(* IEC 61131-3 sources: PortalRobot/Portal_robot/Device/application/FB (part 5) *)

(* ---- FB_ROBOT.st ---- *)
FUNCTION_BLOCK FB_ROBOT
VAR_INPUT
	xUsePhysicalGripperFeedback : BOOL;
	xPhysicalGripperIoReady : BOOL;
	stPhysicalGripperFeedback : ST_GRIPPER_STATUS;
	tPhysicalGripperActionTimeout : TIME := T#10S;
	axMagazineExchangeInProgress : ARRAY [1..2] OF BOOL; // Блокировка адресуется только к меняемому магазину
	xTestInitialize : BOOL;
	auiTestGripperContent : ARRAY [1..2] OF UINT;
	auiTestGripperType : ARRAY [1..2] OF UINT;
	uiTestOrientation : UINT;
	xExternalCommandInhibit : BOOL; // Программный экстренный останов запрещает следующую внешнюю команду
	xSimulationAccelerationEnable : BOOL; // Разрешить ускорение виртуальных таймеров только в симуляции
	uiSimulationTimeFactor : UINT := 1; // Коэффициент виртуального времени 1..100

	stMachine_1_Command : ST_ROBOT_COMMAND; // Команда роботу от первого станка
	stMachine_2_Command : ST_ROBOT_COMMAND; // Команда роботу от второго станка
	stMachine_3_Command : ST_ROBOT_COMMAND; // Команда роботу от третьего станка
	stMagazineCommand   : ST_ROBOT_COMMAND; // Команда роботу от магазина
	stCellCommand       : ST_ROBOT_COMMAND; // Команда позиционирования от менеджера ячейки
	uiBlankPayloadType  : UINT; // Тип заготовки из состояния цикла
	uiDetailPayloadType : UINT; // Тип готовой детали из состояния цикла
	stHmiCommand        : ST_ROBOT_COMMAND; // Ручная команда роботу с HMI
	xReset              : BOOL; // Сброс ошибок робота
	xResetCancel        : BOOL; // Stop/Disable отменяет сброс, не меняя обычную политику останова движения
    xMode               : BOOL; // Режим робота: TRUE — Modbus, FALSE — SoftMotion
	xManual      		: BOOL; // 1 - ручной режим работы, 0 - автоматический режим работы
	xGlobalError        : BOOL; // Глобальная ошибка ячейки
	xEquipmentStopRequired : BOOL; // Владелец оборудования требует зависимую ошибку робота
	ResetDependencies : ST_ROBOT_RESET_DEPENDENCIES; // Снимок отдельных владельцев, только внутренний PLC-контракт
	xModbusBusy         : BOOL; // Внешний робот выполняет команду
	xModbusDone         : BOOL; // Внешний робот завершил команду
	xModbusError        : BOOL; // Ошибка обмена или внешнего робота
	stModbusStatus      : ST_ROBOT_MODBUS_STATUS; // Декодированная обратная связь SC-500
	xHmiDrivesEnable    : BOOL; // Исходный запрос HMI на включение приводов
	xHmiDrivesDisable   : BOOL; // Исходный запрос HMI на отключение приводов
	xHmiStop            : BOOL; // Исходный запрос HMI на остановку
	xHmiDrivesEnableAccepted : BOOL; // RunMotion принял запрос включения в исходном состоянии цикла
	xHmiDrivesDisableAccepted : BOOL; // RunMotion принял запрос отключения в исходном состоянии цикла
	xHmiStopAccepted    : BOOL; // RunMotion принял запрос остановки в исходном состоянии цикла
	xHmiDrivesEnableAllowed : BOOL; // Текущее разрешение включения от владельца Motion-слоя
	xHmiDrivesDisableAllowed : BOOL; // Текущее разрешение отключения от владельца Motion-слоя
	xHmiStopAllowed     : BOOL; // Текущее разрешение остановки от владельца Motion-слоя
	xHmiPermit          : BOOL; // Ручные команды HMI разрешены режимом ячейки
	xManualRecoveryAllowed : BOOL; // Разрешить включение приводов в аварийном ручном восстановлении
	xDrivesPowered      : BOOL; // Все три привода включены
	xDrivesOff          : BOOL; // Все три привода и группа фактически отключены
	xDrivesReady        : BOOL; // Все приводы готовы к движению
	xDriveError         : BOOL; // Активна ошибка оси или группы осей
	xMotionBusy         : BOOL; // Одна из осей выполняет движение
	xMotionResetBusy : BOOL; // Последовательность сброса группы и осей ещё выполняется
	tSoftMotionResetTimeout : TIME := T#30S; // Предел одной принятой попытки сброса
	xSingleAxisMotionBusy : BOOL; // Один из FB_AXIS владеет осью; групповое движение запускать нельзя
	xPointCheckActive : BOOL; // Текущая команда принадлежит проверке сохранённой точки
	xTestAbort : BOOL; // Немедленная отмена активной команды виртуального теста
	rPointCheckSpeedPercent : REAL; // Фактическая скорость проверки 0.1..100 %
	lrGroupAccelerationFactor : LREAL := 1.0; // Общий разгон/торможение групповой траектории, 0.01..1.0
	lrGroupJerkFactor : LREAL := 1.0; // Общий jerk групповой траектории, 0.01..1.0
	tModbusStartTimeout : TIME := T#30S; // Ожидание создания транзакции внешним адаптером
	FaultRequest        : ST_ROBOT_FAULT_REQUEST; // Единый контракт диагностической инъекции
	tGripper1OpenTime   : TIME := T#500MS; // Время открытия первого захвата в модели
	tGripper1CloseTime  : TIME := T#500MS; // Время закрытия первого захвата в модели
	tGripper2OpenTime   : TIME := T#500MS; // Время открытия второго захвата в модели
	tGripper2CloseTime  : TIME := T#500MS; // Время закрытия второго захвата в модели
	tGripperChangeTime  : TIME := T#700MS; // Время смены рабочего захвата в модели

    stPoint : ARRAY [0..GVL_POINT.iPointNumber] OF ST_POINT; // Глобальная таблица точек робота

    xSimBlankAvailable : BOOL; // Начальное наличие заготовки в модели захвата

END_VAR
VAR_OUTPUT
	ResetRecovery : ST_ROBOT_RESET_RECOVERY; // Подтверждение принятой попытки для зависимых владельцев
	GripperCommand : ST_GRIPPER_COMMAND; // Команда для страницы физических выходов
	Command       : ST_ROBOT_COMMAND; // Выбранная команда текущего цикла
	ModbusCommand : ST_ROBOT_COMMAND; // Команда внешнему роботу по Modbus
	Status        : ST_ROBOT_STATUS; // Рабочие статусы робота
	Diag          : ST_ROBOT_DIAG; // Состояние автомата и активная команда
	Error         : ST_ROBOT_ERRORS; // Активные и последние ошибки
	GripperDiag   : ST_GRIPPER_DIAG; // Диагностика внутреннего блока захвата
	GripperError  : ST_GRIPPER_ERRORS; // Активные и последние ошибки захвата
	FaultStatus : ST_ROBOT_FAULT_STATUS; // Сводное состояние инжекторов робота
END_VAR
VAR
	fbMotionManager  : FB_MOTION_MANAGER; // Менеджер перемещения по точкам
    fbGripper        : FB_GRIPPER_SIMULATION; // Модель двухпозиционного захвата
	stGripperCommand : ST_GRIPPER_COMMAND; // Команда внутренней модели захвата

    eState        : E_ROBOT_STATE := E_ROBOT_STATE.IDLE; // Текущее состояние автомата робота
    eActiveAction : E_ROBOT_ACTION := E_ROBOT_ACTION.NONE; // Защёлкнутое действие
    eActivePoint  : E_POINT_NAME; // Защёлкнутая целевая точка
	iActiveSlot   : SINT; // Защёлкнутый слот для всей Modbus-транзакции
	uiActiveMagazineId : UINT; // Защёлкнутый магазин для всей Modbus-транзакции
	uiRobotMagazineContext : UINT; // Физический контекст магазина сохраняется между командами
	xEquipmentStopLatched : BOOL; // Робот остановлен именно аварией обслуживаемого оборудования

	xMotionExecute  : BOOL; // Запрос выполнения перемещения
	xGripperExecute : BOOL; // Запрос выполнения действия захвата
	xManualGripperRequest : BOOL; // Ручной захват разрешён независимо от состояния автомата робота
	xManualGripperOverrideExecute : BOOL; // Прямой импульс FB_GRIPPER из ERROR робота
	eManualGripperAction : E_ROBOT_ACTION; // Действие прямого ручного импульса
	xActiveManualGripper : BOOL; // Текущее действие захвата запущено вручную
	xMagazineCommandActive : BOOL; // Активная команда получена от FB_MAGAZINE
	xMagazineTargetInhibit : BOOL; // Команда входит в магазин, который меняет палеты
	rtReset               : R_TRIG; // Фронт команды сброса робота
	rtHmiDrivesEnable     : R_TRIG; // Фронт запроса включения приводов с HMI
	rtHmiDrivesDisable    : R_TRIG; // Фронт запроса отключения приводов с HMI
	rtHmiStop             : R_TRIG; // Фронт запроса остановки с HMI
	xPowerAllowed         : BOOL; // Визуальная доступность кнопки питания приводов
	xStopAllowed          : BOOL; // Визуальная доступность кнопки остановки
	xResetAllowed         : BOOL; // Визуальная доступность кнопки сброса
	xResetAccepted        : BOOL; // Общий сброс принят владельцем робота
	xExternalResetPending : BOOL; // Удерживает асинхронный Reset до подтверждения SC-500
	xExternalResetIssued  : BOOL; // Reset хотя бы один цикл был передан Modbus-адаптеру
	xSoftMotionResetPending : BOOL; // Один Reset ждёт группу, Motion и захват
	dwResetStopOwners : DWORD; // Владельцы, уже присутствовавшие при принятии Reset
	dwResetLiveCauses : DWORD; // Предыдущий снимок удерживаемых причин этой попытки
	dwResetBusySeen : DWORD; // Владельцы, чей асинхронный сброс действительно запускался
	xEquipmentResetFailed : BOOL; // Новая причина/владелец либо неуспешный терминальный сброс
	tonSoftMotionReset : TON; // Принятая попытка не может оставаться вечной
	xModbusCommandStarted : BOOL; // Текущая команда получила собственную активную транзакцию
	tonModbusStartTimeout : TON; // Защита от вечного ожидания приёма команды адаптером
	fbRobotFaultInjector  : FB_ROBOT_FAULT_INJECTOR; // Безопасная недопустимая команда робота
	xRobotFaultAllowed    : BOOL; // Владелец готов проверить тестовую команду
	uiTestBlankPayloadType : UINT;
	uiTestDetailPayloadType : UINT;
	xTestBlankPayloadPending : BOOL;
	xTestDetailPayloadPending : BOOL;

END_VAR

VAR_IN_OUT
    stMotionManager : ST_MOTION_MANAGER; // Данные менеджера движения
    GroupData       : ST_AXIS_GROUP; // Данные группы осей XYZ
    stPointManager  : ST_POINT_MANAGER; // Данные проверки точки
END_VAR

VAR CONSTANT
	ERR_ROBOT_WRONG_ACTION : DWORD := DWORD#16#0000_0001; // Недопустимое действие робота
    ERR_ROBOT_MOTION       : DWORD := DWORD#16#0000_0002; // Ошибка менеджера движения
    ERR_ROBOT_GRIPPER      : DWORD := DWORD#16#0000_0004; // Ошибка захвата
	ERR_ROBOT_MODBUS_COMM  : DWORD := DWORD#16#0000_0008; // Ошибка связи Modbus TCP
	ERR_ROBOT_STOP         : DWORD := DWORD#16#0000_0010; // Остановка команды робота
	ERR_EXTERNAL_ROBOT     : DWORD := DWORD#16#0000_0020; // Контроллер робота сообщил аварию
	WRN_RESET_EXECUTE_ACTIVE : UINT := 1; // Команда робота ещё активна
	WRN_RESET_STOP_ACTIVE    : UINT := 2; // Команда остановки ещё активна
	WRN_RESET_GLOBAL_ERROR   : UINT := 3; // Глобальная ошибка ещё активна
	WRN_RESET_MOTION_ERROR   : UINT := 4; // Ошибка менеджера движения ещё активна
	WRN_RESET_GRIPPER_ERROR  : UINT := 5; // Ошибка захвата ещё активна
	WRN_RESET_MODBUS_ERROR   : UINT := 6; // Ошибка внешнего робота ещё активна
	WRN_HMI_MANUAL_REQUIRED  : UINT := 7; // Ручная команда запрещена режимом ячейки
	WRN_DRIVES_ENABLE_ERROR  : UINT := 8; // Команда приводов отклонена владельцем Motion-слоя
	WRN_STOP_DRIVES_NOT_READY: UINT := 9; // Остановка недоступна при неготовых приводах
	WRN_SIM_ERROR_NOT_ALLOWED: UINT := 11; // Тестовая команда запрещена текущим состоянием
	WRN_RESET_EQUIPMENT_ERROR : UINT := 18; // WARNING через общий канал: зависимый сброс прерван/не завершён
END_VAR

// --- BEGIN IMPLEMENTATION ---

rtHmiDrivesEnable(CLK := xHmiDrivesEnable);
rtHmiDrivesDisable(CLK := xHmiDrivesDisable);
rtHmiStop(CLK := xHmiStop);

xPowerAllowed := ((NOT xDrivesOff) AND xHmiDrivesDisableAllowed)
	OR (xDrivesOff AND xHmiDrivesEnableAllowed);
xStopAllowed := xHmiStopAllowed;

IF (rtHmiDrivesEnable.Q AND NOT xHmiDrivesEnableAccepted)
OR (rtHmiDrivesDisable.Q AND NOT xHmiDrivesDisableAccepted) THEN
	IF NOT xHmiPermit THEN
		Diag.stWarning.uiCode := WRN_HMI_MANUAL_REQUIRED;
	ELSE
		Diag.stWarning.uiCode := WRN_DRIVES_ENABLE_ERROR;
	END_IF;
	Diag.stWarning.udiSequence := Diag.stWarning.udiSequence + UDINT#1;
	IF Diag.stWarning.udiSequence = UDINT#0 THEN
		Diag.stWarning.udiSequence := UDINT#1;
	END_IF;
END_IF;

IF rtHmiStop.Q
AND NOT xHmiStopAccepted THEN
	IF NOT xHmiPermit THEN
		Diag.stWarning.uiCode := WRN_HMI_MANUAL_REQUIRED;
	ELSE
		Diag.stWarning.uiCode := WRN_STOP_DRIVES_NOT_READY;
	END_IF;
	Diag.stWarning.udiSequence := Diag.stWarning.udiSequence + UDINT#1;
	IF Diag.stWarning.udiSequence = UDINT#0 THEN
		Diag.stWarning.udiSequence := UDINT#1;
	END_IF;
END_IF;

// Команды по умолчанию
xMotionExecute := FALSE;
xGripperExecute := FALSE;
xManualGripperRequest := FALSE;
xManualGripperOverrideExecute := FALSE;
xMagazineCommandActive := FALSE;
xMagazineTargetInhibit := FALSE;

Command.xExecute := FALSE;
Command.xStop := FALSE;
Command.xReset := FALSE;
Command.eAction := E_ROBOT_ACTION.NONE;
Command.eSetPoint := E_POINT_NAME.NONE;
Command.iActiveSlot := 0;
Command.uiMagazineId := UINT#0;

ModbusCommand.xExecute := FALSE;
ModbusCommand.xStop := FALSE;
ModbusCommand.xReset := FALSE;
ModbusCommand.eAction := E_ROBOT_ACTION.NONE;
ModbusCommand.eSetPoint := E_POINT_NAME.NONE;
ModbusCommand.iActiveSlot := 0;
ModbusCommand.uiMagazineId := UINT#0;

//Определяем какой режим работы активен
IF NOT xManual THEN
	IF stCellCommand.xExecute OR stCellCommand.xStop THEN
		Command := stCellCommand;
	ELSIF stMachine_1_Command.xExecute OR stMachine_1_Command.xStop THEN
		Command := stMachine_1_Command;
	ELSIF stMachine_2_Command.xExecute OR stMachine_2_Command.xStop THEN
		Command := stMachine_2_Command;
	ELSIF stMachine_3_Command.xExecute OR stMachine_3_Command.xStop THEN
		Command := stMachine_3_Command;
	ELSIF stMagazineCommand.xExecute OR stMagazineCommand.xStop THEN
		Command := stMagazineCommand;
		xMagazineCommandActive := TRUE;
	END_IF;
ELSE
	IF stMagazineCommand.xExecute OR stMagazineCommand.xStop THEN
		Command := stMagazineCommand;
		xMagazineCommandActive := TRUE;
	ELSE
		Command := stHmiCommand;
	END_IF;
END_IF;

// Смена палет блокирует автоматические команды и операции FB_MAGAZINE
// с этим магазином. Ручная точка HMI не зависит от состояния магазина.
IF (NOT xManual OR xMagazineCommandActive)
AND (Command.uiMagazineId >= UINT#1) AND (Command.uiMagazineId <= UINT#2) THEN
	IF axMagazineExchangeInProgress[Command.uiMagazineId] THEN
		IF (Command.eSetPoint = E_POINT_NAME.MAGAZINE_SAFE)
		OR (Command.eSetPoint = E_POINT_NAME.MAGAZINE_CHANGE)
		OR (Command.eSetPoint = E_POINT_NAME.MAGAZINE_IN_SLOT) THEN
			xMagazineTargetInhibit := TRUE;
		END_IF;
	END_IF;
END_IF;

// Abort теста имеет приоритет над любым владельцем, включая ручную подготовку
// сценария, когда команда ячейки обычно не участвует в выборе.
IF xTestAbort THEN
	Command.xExecute := FALSE;
	Command.xStop := TRUE;
END_IF;

// Уже принятую внешним контроллером команду не прерываем. Запрет действует
// только в IDLE, то есть перед началом следующего высокоуровневого действия.
IF xMode
AND xExternalCommandInhibit
AND (eState = E_ROBOT_STATE.IDLE) THEN
	Command.xExecute := FALSE;
END_IF;

IF xMagazineTargetInhibit AND (eState = E_ROBOT_STATE.IDLE) THEN
	Command.xExecute := FALSE;
END_IF;

// Внешний Stop — самостоятельная приоритетная команда. Он должен дойти до
// адаптера и тогда, когда FB_ROBOT уже защёлкнул ERROR после общей остановки.
IF xMode
AND (xHmiStopAccepted
	OR Command.xStop
	OR (xGlobalError AND stModbusStatus.xBusy)) THEN
	ModbusCommand.xStop := TRUE;
END_IF;

// Класс ошибки определяет оборудование-владелец. FB_ROBOT только выполняет
// зависимую реакцию: активное действие останавливает, неподвижный робот сразу
// переводит в ERROR без бессмысленной команды Stop.
IF xEquipmentStopRequired
AND (eState <> E_ROBOT_STATE.ERROR) THEN
	xEquipmentStopLatched := TRUE;
	IF (eState = E_ROBOT_STATE.MOTION)
	OR (eState = E_ROBOT_STATE.GRIPPER)
	OR (eState = E_ROBOT_STATE.MODBUS) THEN
		Command.xStop := TRUE;
	ELSE
		Error.dwErrorActive := Error.dwErrorActive OR ERR_ROBOT_STOP;
		eState := E_ROBOT_STATE.ERROR;
	END_IF;
END_IF;

// RunRobot уже выполнил все PLC-проверки и передал Execute только принятой
// ручной команде. Захват остаётся независимым от состояния осей и робота.
IF xManual AND stHmiCommand.xExecute THEN
	CASE stHmiCommand.eAction OF
		E_ROBOT_ACTION.UNCLAMP_1,
		E_ROBOT_ACTION.CLAMP_1,
		E_ROBOT_ACTION.UNCLAMP_2,
		E_ROBOT_ACTION.CLAMP_2,
		E_ROBOT_ACTION.ROTATE_TO_BLANK,
		E_ROBOT_ACTION.ROTATE_TO_DETAIL:
			xManualGripperRequest := TRUE;
	END_CASE;
END_IF;

// Готовность сброса рассчитывается после выбора актуального владельца команды.
// Ошибки вложенных FB считаются сбрасываемыми только после снятия удерживаемого
// источника и публикации их собственного xResetAllowed.
rtReset(CLK := xReset);
xResetAllowed := xHmiPermit AND NOT xResetCancel
	AND NOT xTestAbort AND NOT xHmiStop AND NOT xHmiStopAccepted
	AND NOT xSoftMotionResetPending
	AND NOT xExternalResetPending
	AND (NOT xMode OR NOT stModbusStatus.xResetBusy)
	AND (NOT xGlobalError OR xManualRecoveryAllowed)
	AND NOT Command.xExecute
	AND NOT Command.xStop
	AND NOT xMotionBusy
	AND (NOT xMode OR stModbusStatus.xCommunicationAlive)
	AND (xDriveError
		OR (eState = E_ROBOT_STATE.ERROR)
		OR (NOT xMode AND stMotionManager.Status.xError)
		OR (NOT xMode AND fbGripper.Status.xError)
		OR (xMode AND xModbusError))
	AND (xMode OR NOT stMotionManager.Status.xError
		OR FaultStatus.stPoint.xResetAllowed)
	AND (xMode OR NOT fbGripper.Status.xError
		OR FaultStatus.stGripper.xResetAllowed);
xResetAccepted := rtReset.Q AND xResetAllowed;
IF xResetAccepted THEN
	ResetRecovery.udiAttempt := ResetRecovery.udiAttempt + UDINT#1;
	IF ResetRecovery.udiAttempt = UDINT#0 THEN ResetRecovery.udiAttempt := UDINT#1; END_IF;
	dwResetStopOwners := ResetDependencies.dwStopOwners;
	dwResetLiveCauses := ResetDependencies.dwLiveCauses;
	dwResetBusySeen := ResetDependencies.dwResetBusy;
END_IF;
xEquipmentResetFailed := FALSE;
IF (xSoftMotionResetPending OR xExternalResetPending) AND NOT xResetAccepted THEN
	// Нового владельца или повторный фронт физической причины нельзя принять
	// за хвост старого сброса. Падение Busy само по себе успехом не является.
	xEquipmentResetFailed := ((ResetDependencies.dwStopOwners AND NOT dwResetStopOwners) <> DWORD#0)
		OR ((ResetDependencies.dwLiveCauses AND NOT dwResetLiveCauses) <> DWORD#0)
		OR ((dwResetBusySeen AND NOT ResetDependencies.dwResetBusy
			AND ResetDependencies.dwStopOwners) <> DWORD#0);
	dwResetLiveCauses := ResetDependencies.dwLiveCauses;
	dwResetBusySeen := dwResetBusySeen OR ResetDependencies.dwResetBusy;
END_IF;
// Общий Reset запускает Motion-сброс раньше FB_ROBOT. Если группа была в
// ErrorStop, одноцикловый импульс уже закончится к моменту её восстановления;
// защёлкиваем намерение оператора до исчезновения первичной Motion-ошибки.
IF xMode THEN
	xSoftMotionResetPending := FALSE;
ELSIF xResetAccepted
AND (eState = E_ROBOT_STATE.ERROR) THEN
	xSoftMotionResetPending := TRUE;
END_IF;
IF xMode AND xResetAccepted THEN
	xExternalResetPending := TRUE;
	xExternalResetIssued := FALSE;
ELSIF NOT xMode THEN
	xExternalResetPending := FALSE;
	xExternalResetIssued := FALSE;
END_IF;

tonSoftMotionReset(IN := xSoftMotionResetPending OR xExternalResetPending, PT := tSoftMotionResetTimeout);
IF xSoftMotionResetPending AND NOT xResetAccepted
AND (tonSoftMotionReset.Q
	OR xEquipmentResetFailed OR xResetCancel
	OR xTestAbort OR NOT xHmiPermit OR Command.xExecute OR Command.xStop OR xHmiStop OR xHmiStopAccepted
	OR (xGlobalError AND NOT xManualRecoveryAllowed)
	OR (xDriveError AND NOT xMotionResetBusy)
	OR (fbGripper.Status.xError AND NOT FaultStatus.stGripper.xResetAllowed)
	OR (stMotionManager.Status.xError AND NOT FaultStatus.stPoint.xResetAllowed)) THEN
	xSoftMotionResetPending := FALSE;
	IF xEquipmentResetFailed OR (tonSoftMotionReset.Q AND xEquipmentStopRequired) THEN
		Diag.stWarning.uiCode := WRN_RESET_EQUIPMENT_ERROR;
	ELSIF fbGripper.Status.xError THEN
		Diag.stWarning.uiCode := WRN_RESET_GRIPPER_ERROR;
	ELSE
		Diag.stWarning.uiCode := WRN_RESET_MOTION_ERROR;
	END_IF;
	Diag.stWarning.udiSequence := Diag.stWarning.udiSequence + UDINT#1;
	IF Diag.stWarning.udiSequence = UDINT#0 THEN Diag.stWarning.udiSequence := UDINT#1; END_IF;
END_IF;

// После неуспешной попытки адаптер публикует явный результат. Снимаем уровень,
// чтобы следующее осознанное нажатие Reset снова дошло до его R_TRIG.
IF xExternalResetPending AND xExternalResetIssued AND NOT xResetAccepted
AND (stModbusStatus.xResetFailed OR NOT stModbusStatus.xCommunicationAlive
	OR tonSoftMotionReset.Q OR xEquipmentResetFailed OR xResetCancel
	OR xTestAbort OR Command.xStop OR xHmiStop OR xHmiStopAccepted OR NOT xHmiPermit
	OR (xGlobalError AND NOT xManualRecoveryAllowed)) THEN
	xExternalResetPending := FALSE;
	xExternalResetIssued := FALSE;
	IF xEquipmentResetFailed OR (tonSoftMotionReset.Q AND xEquipmentStopRequired) THEN
		Diag.stWarning.uiCode := WRN_RESET_EQUIPMENT_ERROR;
	ELSE
		Diag.stWarning.uiCode := WRN_RESET_MODBUS_ERROR;
	END_IF;
	Diag.stWarning.udiSequence := Diag.stWarning.udiSequence + UDINT#1;
	IF Diag.stWarning.udiSequence = UDINT#0 THEN Diag.stWarning.udiSequence := UDINT#1; END_IF;
END_IF;

// Недопустимое действие проверяется в IDLE до запуска Motion или захвата.
xRobotFaultAllowed := (eState = E_ROBOT_STATE.IDLE)
	AND NOT Command.xExecute
	AND NOT Command.xStop
	AND NOT xMode
	AND NOT xGlobalError
	AND NOT xDriveError
	AND (Error.dwErrorActive = DWORD#0)
	AND NOT stMotionManager.Status.xError
	AND NOT fbGripper.Status.xError;

fbRobotFaultInjector(
	Request := FaultRequest,
	xOwnerAllowed := xRobotFaultAllowed
);
FaultStatus.stRobot := fbRobotFaultInjector.Status;

IF fbRobotFaultInjector.Status.xRejected THEN
	Diag.stWarning.uiCode := WRN_SIM_ERROR_NOT_ALLOWED;
	Diag.stWarning.udiSequence := Diag.stWarning.udiSequence + UDINT#1;
	IF Diag.stWarning.udiSequence = UDINT#0 THEN
		Diag.stWarning.udiSequence := UDINT#1;
	END_IF;
END_IF;

IF fbRobotFaultInjector.xWrongAction THEN
	Command.xExecute := TRUE;
	Command.xStop := FALSE;
	Command.eAction := E_ROBOT_ACTION.NONE;
	Command.eSetPoint := E_POINT_NAME.NONE;
END_IF;

Command.xReset := xResetAccepted;

IF rtReset.Q
AND ((eState = E_ROBOT_STATE.ERROR) OR xDriveError)
AND NOT xResetAccepted THEN
	IF NOT xHmiPermit THEN
		Diag.stWarning.uiCode := WRN_HMI_MANUAL_REQUIRED;
	ELSIF eState <> E_ROBOT_STATE.ERROR THEN
		// Ошибку Motion-слоя сбрасывают оси и группа тем же общим импульсом.
		Diag.stWarning.uiCode := UINT#0;
    ELSIF Command.xExecute THEN
        Diag.stWarning.uiCode := WRN_RESET_EXECUTE_ACTIVE;
    ELSIF Command.xStop THEN
        Diag.stWarning.uiCode := WRN_RESET_STOP_ACTIVE;
    ELSIF xGlobalError AND NOT xManualRecoveryAllowed THEN
        Diag.stWarning.uiCode := WRN_RESET_GLOBAL_ERROR;
    ELSIF stMotionManager.Status.xError
	OR (NOT xMode AND xDriveError) THEN
        Diag.stWarning.uiCode := WRN_RESET_MOTION_ERROR;
    ELSIF fbGripper.Status.xError THEN
        Diag.stWarning.uiCode := WRN_RESET_GRIPPER_ERROR;
    ELSIF xModbusError THEN
        Diag.stWarning.uiCode := WRN_RESET_MODBUS_ERROR;
    ELSE
        Diag.stWarning.uiCode := UINT#0;
    END_IF;

    IF Diag.stWarning.uiCode <> UINT#0 THEN
        Diag.stWarning.udiSequence := Diag.stWarning.udiSequence + UDINT#1;
        IF Diag.stWarning.udiSequence = UDINT#0 THEN
            Diag.stWarning.udiSequence := UDINT#1;
        END_IF;
    END_IF;
END_IF;

// =====================================================
// Автомат FB_ROBOT
// =====================================================

// Таймаут исполнения принадлежит FB_ROBOT_MODBUS, но до создания активной
// транзакции его TON ещё не работает. Отдельно ограничиваем фазу ожидания Busy.
tonModbusStartTimeout(
	IN := xMode
		AND (eState = E_ROBOT_STATE.MODBUS)
		AND NOT xModbusCommandStarted,
	PT := tModbusStartTimeout
);

// Ошибка оси или группы является первопричиной в Motion-слое и отдельной
// каскадной ошибкой робота для его публичного статуса и журнала.
IF NOT xMode AND xDriveError THEN
	Error.dwErrorActive := Error.dwErrorActive OR ERR_ROBOT_MOTION;
	eState := E_ROBOT_STATE.ERROR;
ELSIF NOT xMode AND stMotionManager.Status.xError THEN
	// Отмена задания при ручном I/O не скрывает аварию вложенного владельца.
	Error.dwErrorActive := Error.dwErrorActive OR ERR_ROBOT_MOTION;
	eState := E_ROBOT_STATE.ERROR;
ELSIF NOT xMode AND fbGripper.Status.xError THEN
	Error.dwErrorActive := Error.dwErrorActive OR ERR_ROBOT_GRIPPER;
	eState := E_ROBOT_STATE.ERROR;
ELSIF xMode AND xModbusError THEN
	IF stModbusStatus.xRobotAlarm THEN
		Error.dwErrorActive := Error.dwErrorActive OR ERR_EXTERNAL_ROBOT;
	ELSE
		Error.dwErrorActive := Error.dwErrorActive OR ERR_ROBOT_MODBUS_COMM;
	END_IF;
	eState := E_ROBOT_STATE.ERROR;
END_IF;

CASE eState OF

    E_ROBOT_STATE.IDLE:

        Status.xBusy := FALSE;
        Status.xDone := FALSE;
        Status.xError := FALSE;

        IF Command.xExecute THEN
            eActiveAction := Command.eAction;
            eActivePoint := Command.eSetPoint;
			iActiveSlot := Command.iActiveSlot;
			uiActiveMagazineId := Command.uiMagazineId;
			IF (Command.uiMagazineId >= UINT#1)
			AND (Command.uiMagazineId <= UINT#2)
			AND (Command.eAction = E_ROBOT_ACTION.MOVE_TO_POINT)
			AND ((Command.eSetPoint = E_POINT_NAME.MAGAZINE_IN_SLOT)
				OR (Command.eSetPoint = E_POINT_NAME.MAGAZINE_CHANGE)) THEN
				uiRobotMagazineContext := Command.uiMagazineId;
			END_IF;

            IF xMode THEN
				xModbusCommandStarted := FALSE;
				eState := E_ROBOT_STATE.MODBUS;

            ELSE
                CASE Command.eAction OF

                    E_ROBOT_ACTION.MOVE_TO_POINT:
                        // CODESYS переводит группу в ошибку, если GroupMoving
                        // запускается при активном single-axis FB. Команда
                        // остаётся в IDLE до освобождения всех FB_AXIS.
                        IF xDrivesReady AND NOT xMotionBusy THEN
                            eState := E_ROBOT_STATE.MOTION;
                        END_IF;

                    E_ROBOT_ACTION.UNCLAMP_1,
                    E_ROBOT_ACTION.CLAMP_1,
                    E_ROBOT_ACTION.UNCLAMP_2,
                    E_ROBOT_ACTION.CLAMP_2,
                    E_ROBOT_ACTION.ROTATE_TO_BLANK,
                    E_ROBOT_ACTION.ROTATE_TO_DETAIL:
						xActiveManualGripper := xManualGripperRequest;
                        eState := E_ROBOT_STATE.GRIPPER;

                ELSE
                    Error.dwErrorActive :=
                        Error.dwErrorActive OR ERR_ROBOT_WRONG_ACTION;

                    eState := E_ROBOT_STATE.ERROR;
                END_CASE;
            END_IF;
        END_IF;

    E_ROBOT_STATE.MOTION:

        Status.xBusy := TRUE;
        xMotionExecute := NOT xSingleAxisMotionBusy;

		IF xHmiStopAccepted OR Command.xStop THEN
			// Операторский Stop отменяет действие штатно. Stop от оборудования
			// дополнительно защёлкивает зависимую ошибку робота.
            xMotionExecute := FALSE;
            Status.xBusy := FALSE;
            Status.xDone := FALSE;
            eActiveAction := E_ROBOT_ACTION.NONE;
            eActivePoint := E_POINT_NAME.NONE;
			IF xEquipmentStopRequired THEN
				Error.dwErrorActive := Error.dwErrorActive OR ERR_ROBOT_STOP;
				eState := E_ROBOT_STATE.ERROR;
			ELSE
				eState := E_ROBOT_STATE.IDLE;
			END_IF;

        ELSIF xGlobalError THEN
            Error.dwErrorActive := Error.dwErrorActive OR ERR_ROBOT_STOP;
            eState := E_ROBOT_STATE.ERROR;

        ELSIF stMotionManager.Status.xError THEN
            Error.dwErrorActive := Error.dwErrorActive OR ERR_ROBOT_MOTION;
            eState := E_ROBOT_STATE.ERROR;

		ELSIF stMotionManager.Status.xDone THEN
			IF (eActiveAction = E_ROBOT_ACTION.MOVE_TO_POINT)
			AND (eActivePoint <> E_POINT_NAME.MAGAZINE_IN_SLOT)
			AND (eActivePoint <> E_POINT_NAME.MAGAZINE_CHANGE) THEN
				uiRobotMagazineContext := UINT#0;
			END_IF;
            eState := E_ROBOT_STATE.DONE;
        END_IF;

	E_ROBOT_STATE.GRIPPER:

        Status.xBusy := TRUE;
        xGripperExecute := TRUE;

		IF xTestAbort THEN
			xGripperExecute := FALSE;
			Status.xBusy := FALSE;
			Status.xDone := FALSE;
			xActiveManualGripper := FALSE;
			eActiveAction := E_ROBOT_ACTION.NONE;
			eActivePoint := E_POINT_NAME.NONE;
			eState := E_ROBOT_STATE.IDLE;

		ELSIF xEquipmentStopRequired THEN
			xGripperExecute := FALSE;
			Error.dwErrorActive := Error.dwErrorActive OR ERR_ROBOT_STOP;
			eState := E_ROBOT_STATE.ERROR;

		ELSIF xGlobalError AND NOT xActiveManualGripper THEN
            Error.dwErrorActive := Error.dwErrorActive OR ERR_ROBOT_STOP;
            eState := E_ROBOT_STATE.ERROR;

        ELSIF fbGripper.Status.xError THEN
            Error.dwErrorActive := Error.dwErrorActive OR ERR_ROBOT_GRIPPER;
            eState := E_ROBOT_STATE.ERROR;

        ELSIF fbGripper.Status.xDone THEN
			xActiveManualGripper := FALSE;
            eState := E_ROBOT_STATE.DONE;
        END_IF;

	E_ROBOT_STATE.DONE:

        Status.xBusy := FALSE;
        Status.xDone := TRUE;

        IF NOT xMode THEN
        CASE eActiveAction OF

            E_ROBOT_ACTION.MOVE_TO_POINT:
                xMotionExecute := TRUE;

            E_ROBOT_ACTION.UNCLAMP_1,
            E_ROBOT_ACTION.CLAMP_1,
            E_ROBOT_ACTION.UNCLAMP_2,
            E_ROBOT_ACTION.CLAMP_2,
            E_ROBOT_ACTION.ROTATE_TO_BLANK,
            E_ROBOT_ACTION.ROTATE_TO_DETAIL:
                xGripperExecute := TRUE;

        END_CASE;
        END_IF;

		IF NOT Command.xExecute THEN
			// Владелец уже снял Execute: в этом же цикле погасить запрос
			// вложенному FB до очистки action/point. Иначе при быстром
			// SoftMotion движении один скан уходил как Execute=TRUE + point=NONE,
			// а FB_MOTION_MANAGER закономерно валил нулевую точку.
			xMotionExecute := FALSE;
			xGripperExecute := FALSE;
            Status.xDone := FALSE;
			xModbusCommandStarted := FALSE;
            eActiveAction := E_ROBOT_ACTION.NONE;
			eActivePoint := E_POINT_NAME.NONE;
			iActiveSlot := SINT#0;
			uiActiveMagazineId := UINT#0;
			eState := E_ROBOT_STATE.IDLE;
        END_IF;

	E_ROBOT_STATE.MODBUS:
		Status.xBusy := TRUE;
		// Execute — импульс от владельца команды. Адаптер Modbus может
		// быть занят FC03/FC16 дольше этого импульса. Поэтому до терминального
		// ответа передаём защёлкнутые action/point/slot, а не уже снятый Command.
		ModbusCommand.xExecute := TRUE;
		ModbusCommand.eAction := eActiveAction;
		ModbusCommand.eSetPoint := eActivePoint;
		ModbusCommand.iActiveSlot := iActiveSlot;
		ModbusCommand.uiMagazineId := uiActiveMagazineId;
		IF xModbusBusy THEN
			xModbusCommandStarted := TRUE;
		END_IF;

		IF xTestAbort THEN
			ModbusCommand.xStop := TRUE;
			IF NOT stModbusStatus.xBusy THEN
				Status.xBusy := FALSE;
				Status.xDone := FALSE;
				xModbusCommandStarted := FALSE;
				eActiveAction := E_ROBOT_ACTION.NONE;
				eActivePoint := E_POINT_NAME.NONE;
				iActiveSlot := SINT#0;
				uiActiveMagazineId := UINT#0;
				eState := E_ROBOT_STATE.IDLE;
			END_IF;
		ELSIF Command.xStop OR xHmiStopAccepted OR xGlobalError THEN
			ModbusCommand.xStop := TRUE;
			Error.dwErrorActive := Error.dwErrorActive OR ERR_ROBOT_STOP;
			eState := E_ROBOT_STATE.ERROR;
		ELSIF xModbusError THEN
			IF stModbusStatus.xRobotAlarm THEN
				Error.dwErrorActive := Error.dwErrorActive OR ERR_EXTERNAL_ROBOT;
			ELSE
				Error.dwErrorActive := Error.dwErrorActive OR ERR_ROBOT_MODBUS_COMM;
			END_IF;
			eState := E_ROBOT_STATE.ERROR;
		ELSIF tonModbusStartTimeout.Q THEN
			// Адаптер не создал собственную транзакцию: не оставляем публичный
			// xBusy висеть бесконечно без CommandSeq и физического движения.
			ModbusCommand.xExecute := FALSE;
			Error.dwErrorActive := Error.dwErrorActive OR ERR_ROBOT_MODBUS_COMM;
			eState := E_ROBOT_STATE.ERROR;
		ELSIF xModbusCommandStarted AND xModbusDone THEN
			IF (eActiveAction = E_ROBOT_ACTION.MOVE_TO_POINT)
			AND (eActivePoint <> E_POINT_NAME.MAGAZINE_IN_SLOT)
			AND (eActivePoint <> E_POINT_NAME.MAGAZINE_CHANGE) THEN
				uiRobotMagazineContext := UINT#0;
			END_IF;
			eState := E_ROBOT_STATE.DONE;
		END_IF;

    E_ROBOT_STATE.ERROR:

        Status.xBusy := FALSE;
        Status.xDone := FALSE;
        Status.xError := TRUE;

		// Ошибка координатного робота не блокирует независимый ручной захват.
		// Собственная ошибка FB_GRIPPER по-прежнему требует штатного сброса.
		IF NOT xMode AND xManualGripperRequest AND NOT fbGripper.Status.xError THEN
			xManualGripperOverrideExecute := TRUE;
			eManualGripperAction := stHmiCommand.eAction;
		END_IF;

		// В Modbus-режиме входной Reset только защёлкивает запрос для адаптера.
		// Локальную ошибку можно снять лишь после подтверждённого исчезновения
		// внешней аварии; иначе xExternalResetPending очистится до записи 1004.
		IF ((NOT xMode AND (xResetAccepted OR xSoftMotionResetPending))
			OR (xMode
				AND xExternalResetPending
				AND xExternalResetIssued
				AND stModbusStatus.xResetDone
				AND NOT xModbusError
				AND NOT stModbusStatus.xBusy
				AND (stModbusStatus.uiExecutionState =
					TO_UINT(E_ROBOT_MODBUS_EXECUTION_STATE.IDLE))))
        AND NOT Command.xExecute
        AND NOT Command.xStop
        AND NOT xEquipmentStopRequired
        AND (NOT xGlobalError OR xManualRecoveryAllowed)
		AND (xMode OR NOT stMotionManager.Status.xError)
		AND (xMode OR NOT xDriveError)
		AND (xMode OR NOT xMotionResetBusy)
		AND (xMode OR NOT fbGripper.Status.xError)
		AND (NOT xMode OR stModbusStatus.xCommunicationAlive) THEN

			Error.dwErrorLast := Error.dwErrorActive;
			Error.dwErrorActive := DWORD#0;
            Status.xError := FALSE;
			xExternalResetPending := FALSE;
			xExternalResetIssued := FALSE;
			xSoftMotionResetPending := FALSE;
			xModbusCommandStarted := FALSE;
			xActiveManualGripper := FALSE;
			xEquipmentStopLatched := FALSE;
            eActiveAction := E_ROBOT_ACTION.NONE;
			eActivePoint := E_POINT_NAME.NONE;
			iActiveSlot := SINT#0;
			uiActiveMagazineId := UINT#0;
			eState := E_ROBOT_STATE.IDLE;
        END_IF;

END_CASE;

IF xMode AND xExternalResetPending THEN
	ModbusCommand.xReset := TRUE;
	xExternalResetIssued := TRUE;
END_IF;

// =====================================================
// Формирование команды FB_MOTION_MANAGER
// =====================================================

stMotionManager.Command.xExecute := NOT xMode AND xMotionExecute;
stMotionManager.Command.eTargetPoint := eActivePoint;
stMotionManager.Command.xReset := NOT xMode AND xResetAccepted;
stMotionManager.Command.xStop := NOT xMode AND (xHmiStopAccepted OR Command.xStop);
stMotionManager.Command.xGlobalError :=
    (NOT xMode AND xGlobalError AND NOT xManualRecoveryAllowed);

// =====================================================
// Вызов FB_MOTION_MANAGER
// =====================================================

fbMotionManager(
    stPoint := stPoint,
    xReset := NOT xMode AND xResetAccepted,
	FaultRequest := FaultRequest.stPoint,
	xSpeedFactorOverride := xPointCheckActive,
	lrSpeedFactorOverride := REAL_TO_LREAL(rPointCheckSpeedPercent) / 100.0,
	lrAccelerationFactor := lrGroupAccelerationFactor,
	lrJerkFactor := lrGroupJerkFactor,
    stMotionManager := stMotionManager,
    GroupData := GroupData,
    stPointManager := stPointManager
);
FaultStatus.stPoint := fbMotionManager.FaultStatus;

// =====================================================
// Вызов FB_GRIPPER
// =====================================================

stGripperCommand.xExecute := NOT xMode
	AND (xGripperExecute OR xManualGripperOverrideExecute);
stGripperCommand.xReset := NOT xMode AND xResetAccepted;
stGripperCommand.xGripper1Open := fbGripper.Status.xGripper1Open;
stGripperCommand.xGripper2Open := fbGripper.Status.xGripper2Open;
stGripperCommand.xRotateToDetail := fbGripper.Status.xRotatedToDetail;
IF xManualGripperOverrideExecute THEN
	stGripperCommand.eAction := eManualGripperAction;
ELSE
	stGripperCommand.eAction := eActiveAction;
END_IF;
CASE stGripperCommand.eAction OF
	E_ROBOT_ACTION.UNCLAMP_1: stGripperCommand.xGripper1Open := TRUE;
	E_ROBOT_ACTION.CLAMP_1: stGripperCommand.xGripper1Open := FALSE;
	E_ROBOT_ACTION.UNCLAMP_2: stGripperCommand.xGripper2Open := TRUE;
	E_ROBOT_ACTION.CLAMP_2: stGripperCommand.xGripper2Open := FALSE;
	E_ROBOT_ACTION.ROTATE_TO_BLANK: stGripperCommand.xRotateToDetail := FALSE;
	E_ROBOT_ACTION.ROTATE_TO_DETAIL: stGripperCommand.xRotateToDetail := TRUE;
END_CASE;

GripperCommand := stGripperCommand;
fbGripper(
	xUsePhysicalFeedback := xUsePhysicalGripperFeedback AND NOT xMode,
	xPhysicalIoReady := xPhysicalGripperIoReady,
	PhysicalFeedback := stPhysicalGripperFeedback,
	tPhysicalActionTimeout := tPhysicalGripperActionTimeout,
	// Положение и захваты робота не подменяются записью сценария: runner
	// приводит их в нужное состояние штатными командами.
	xTestInitialize := FALSE,
	auiTestContent := auiTestGripperContent,
	uiTestOrientation := uiTestOrientation,
	Command := stGripperCommand,
	FaultRequest := FaultRequest.stGripper,
	xSimulationAccelerationEnable := xSimulationAccelerationEnable,
	uiSimulationTimeFactor := uiSimulationTimeFactor,
	tGripper1OpenTime := tGripper1OpenTime,
	tGripper1CloseTime := tGripper1CloseTime,
	tGripper2OpenTime := tGripper2OpenTime,
	tGripper2CloseTime := tGripper2CloseTime,
	tRotateTime := tGripperChangeTime,
	Diag => GripperDiag,
	Error => GripperError
);
FaultStatus.stGripper := fbGripper.FaultStatus;

IF xTestInitialize THEN
	uiTestBlankPayloadType := auiTestGripperType[1];
	uiTestDetailPayloadType := auiTestGripperType[2];
	xTestBlankPayloadPending := auiTestGripperContent[1] = UINT#1;
	xTestDetailPayloadPending := auiTestGripperContent[2] = UINT#2;
	uiRobotMagazineContext := UINT#0;
	xEquipmentStopLatched := FALSE;
	xSoftMotionResetPending := FALSE;
END_IF;

// =====================================================
// Общие статусы
// =====================================================

IF xMode THEN
	CASE stModbusStatus.uiCurrentPoint OF
		10: Status.eCurrentPoint := E_POINT_NAME.MACHINE_1_ABOVE;
		11: Status.eCurrentPoint := E_POINT_NAME.MACHINE_1_INSIDE;
		12: Status.eCurrentPoint := E_POINT_NAME.MACHINE_1_CHUCK_APROACH;
		13: Status.eCurrentPoint := E_POINT_NAME.MACHINE_1_CHUCK_POSITION;
		14: Status.eCurrentPoint := E_POINT_NAME.MACHINE_2_ABOVE;
		15: Status.eCurrentPoint := E_POINT_NAME.MACHINE_2_INSIDE;
		16: Status.eCurrentPoint := E_POINT_NAME.MACHINE_2_CHUCK_APROACH;
		17: Status.eCurrentPoint := E_POINT_NAME.MACHINE_2_CHUCK_POSITION;
		18: Status.eCurrentPoint := E_POINT_NAME.MACHINE_3_ABOVE;
		19: Status.eCurrentPoint := E_POINT_NAME.MACHINE_3_INSIDE;
		20: Status.eCurrentPoint := E_POINT_NAME.MACHINE_3_CHUCK_APROACH;
		21: Status.eCurrentPoint := E_POINT_NAME.MACHINE_3_CHUCK_POSITION;
		22: Status.eCurrentPoint := E_POINT_NAME.HOME_SAFETY;
		23: Status.eCurrentPoint := E_POINT_NAME.MAGAZINE_SAFE;
		24: Status.eCurrentPoint := E_POINT_NAME.MAGAZINE_CHANGE;
		25: Status.eCurrentPoint := E_POINT_NAME.MAGAZINE_IN_SLOT;
	ELSE
		Status.eCurrentPoint := E_POINT_NAME.NONE;
	END_CASE;
	Status.xGripper1Open := (stModbusStatus.uiGripperStatus AND UINT#16#0001) <> UINT#0;
	Status.xGripper1Closed := (stModbusStatus.uiGripperStatus AND UINT#16#0002) <> UINT#0;
	Status.xGripper2Open := (stModbusStatus.uiGripperStatus AND UINT#16#0004) <> UINT#0;
	Status.xGripper2Closed := (stModbusStatus.uiGripperStatus AND UINT#16#0008) <> UINT#0;
	Status.xRotatedToBlank := (stModbusStatus.uiGripperStatus AND UINT#16#0010) <> UINT#0;
	Status.xRotatedToDetail := (stModbusStatus.uiGripperStatus AND UINT#16#0020) <> UINT#0;
ELSE
	Status.eCurrentPoint := stMotionManager.Status.eCurrentPoint;
	Status.xGripper1Open := fbGripper.Status.xGripper1Open;
	Status.xGripper1Closed := fbGripper.Status.xGripper1Closed;
	Status.xGripper2Open := fbGripper.Status.xGripper2Open;
	Status.xGripper2Closed := fbGripper.Status.xGripper2Closed;
	Status.xRotatedToBlank := fbGripper.Status.xRotatedToBlank;
	Status.xRotatedToDetail := fbGripper.Status.xRotatedToDetail;
END_IF;

Status.xBlankAvailable := Status.xGripper1Closed;
Status.xDetailAvailable := Status.xGripper2Closed;
IF Status.xGripper1Open THEN
	Status.uiBlankPayloadType := UINT#0;
	IF NOT xTestBlankPayloadPending THEN
		uiTestBlankPayloadType := UINT#0;
	END_IF;
ELSIF Status.xGripper1Closed THEN
	// Во время загрузки тестового сценария его тип относится к уже заданному
	// содержимому захвата и имеет приоритет над метаданными предыдущего цикла.
	IF xTestBlankPayloadPending
	AND (uiTestBlankPayloadType >= UINT#1)
	AND (uiTestBlankPayloadType <= UINT#3) THEN
		Status.uiBlankPayloadType := uiTestBlankPayloadType;
	ELSIF (uiBlankPayloadType >= UINT#1) AND (uiBlankPayloadType <= UINT#3) THEN
		Status.uiBlankPayloadType := uiBlankPayloadType;
		uiTestBlankPayloadType := uiBlankPayloadType;
	ELSIF (uiTestBlankPayloadType >= UINT#1)
	AND (uiTestBlankPayloadType <= UINT#3) THEN
		Status.uiBlankPayloadType := uiTestBlankPayloadType;
	ELSE
		Status.uiBlankPayloadType := UINT#0;
	END_IF;
	xTestBlankPayloadPending := FALSE;
END_IF;
IF Status.xGripper2Open THEN
	Status.uiDetailPayloadType := UINT#0;
	IF NOT xTestDetailPayloadPending THEN
		uiTestDetailPayloadType := UINT#0;
	END_IF;
ELSIF Status.xGripper2Closed THEN
	IF xTestDetailPayloadPending
	AND (uiTestDetailPayloadType >= UINT#1)
	AND (uiTestDetailPayloadType <= UINT#3) THEN
		Status.uiDetailPayloadType := uiTestDetailPayloadType;
	ELSIF (uiDetailPayloadType >= UINT#1) AND (uiDetailPayloadType <= UINT#3) THEN
		Status.uiDetailPayloadType := uiDetailPayloadType;
		uiTestDetailPayloadType := uiDetailPayloadType;
	ELSIF (uiTestDetailPayloadType >= UINT#1)
	AND (uiTestDetailPayloadType <= UINT#3) THEN
		Status.uiDetailPayloadType := uiTestDetailPayloadType;
	ELSE
		Status.uiDetailPayloadType := UINT#0;
	END_IF;
	xTestDetailPayloadPending := FALSE;
END_IF;
Status.xPowerAllowed := xPowerAllowed;
Status.xStopAllowed := xStopAllowed;
Status.xResetAllowed := xResetAllowed;
ResetRecovery.xActive := xSoftMotionResetPending OR xExternalResetPending;
// Положительное подтверждение относится только к первичным зависимостям.
// Родитель остаётся в ERROR, пока оборудование снимает свой старый каскад.
ResetRecovery.xDependenciesReady := ResetRecovery.xActive
	AND xHmiPermit AND NOT xResetCancel AND NOT xTestAbort AND NOT Command.xExecute AND NOT Command.xStop
	AND NOT xHmiStop AND NOT xHmiStopAccepted AND NOT xMotionBusy
	AND (NOT xGlobalError OR xManualRecoveryAllowed)
	AND ((NOT xMode AND NOT xDriveError AND NOT xMotionResetBusy
		AND NOT stMotionManager.Status.xError AND NOT fbGripper.Status.xError)
		OR (xMode AND xExternalResetIssued AND stModbusStatus.xResetDone
			AND NOT xModbusError AND stModbusStatus.xCommunicationAlive
			AND NOT stModbusStatus.xBusy
			AND (stModbusStatus.uiExecutionState = TO_UINT(E_ROBOT_MODBUS_EXECUTION_STATE.IDLE))));
Status.uiMagazineContext := uiRobotMagazineContext;

Diag.eState := eState;
Diag.eActiveAction := eActiveAction;
Diag.eActivePoint := eActivePoint;
Error.dwAlarmActive := Error.dwErrorActive;
Status.xExternalError := ((Error.dwErrorActive AND (ERR_ROBOT_MOTION OR ERR_ROBOT_GRIPPER)) <> DWORD#0)
	OR xEquipmentStopLatched;

IF Error.dwErrorActive <> DWORD#0 THEN
	Error.dwErrorLast := Error.dwErrorActive;
END_IF;

Error.stErrorActive := UpdateErrorView(dwError := Error.dwErrorActive);
Error.stErrorLast := UpdateErrorView(dwError := Error.dwErrorLast);
FaultStatus.stRobot.xResetAllowed := Status.xResetAllowed
	AND NOT FaultStatus.stRobot.xBusy;

(* ---- FB_ROBOT_MODBUS.st ---- *)
{attribute 'no_assign'}
FUNCTION_BLOCK FB_ROBOT_MODBUS
VAR_INPUT
	xEnable          : BOOL; // Применён режим MODBUS_TCP
	xReconnect       : BOOL; // Настройки изменены, выполнить reconnect
	Config           : ST_ROBOT_MODBUS_CONFIG;
	Command          : ST_ROBOT_COMMAND; // Семантическая команда FB_ROBOT
END_VAR
VAR_OUTPUT
	Status           : ST_ROBOT_MODBUS_STATUS;
END_VAR
VAR_IN_OUT
	auiWriteRegisters : ARRAY [0..8] OF UINT; // Документные адреса 1001..1009
	auiReadRegisters  : ARRAY [0..16] OF UINT; // Документные адреса 1101..1117
END_VAR
VAR
	{attribute 'no_assign'}
	fbClient       : ModbusFB.ClientTCP;
	fbRead         : ModbusFB.ClientRequestReadHoldingRegisters;
	fbWrite        : ModbusFB.ClientRequestWriteMultipleRegisters;
	eState         : E_ROBOT_MODBUS_CLIENT_STATE := E_ROBOT_MODBUS_CLIENT_STATE.DISABLED;
	xConnect       : BOOL;
	xReadExecute   : BOOL;
	xWriteExecute  : BOOL;
	xStatusFresh   : BOOL;
	xCommandArmed  : BOOL;
	xCommandActive : BOOL;
	xWritePending  : BOOL;
	xHeartbeatChanged : BOOL;
	xHeartbeatSeen : BOOL;
	xPlcHeartbeatDue : BOOL;
	xStopPending   : BOOL;
	xResetPending  : BOOL;
	xResetInProgress : BOOL;
	xResetWriteDone : BOOL; // FC16 с Reset=1 подтверждена сервером
	tonResetAttempt : TON;
	xControlClearPending : BOOL;
	rtStop         : R_TRIG;
	rtReset        : R_TRIG;
	rtReconnect    : R_TRIG;
	tonPoll        : TON;
	tonPlcHeartbeat: TON;
	tonRobotHeartbeat : TON;
	tonCommunicationGrace : TON;
	tonCommandTimeout : TON;
	tonReconnect   : TON;
	uiCommandSeq   : UINT;
	uiActiveSeq    : UINT;
	uiDecodedRobotHeartbeat : UINT; // Heartbeat из последнего завершённого FC03
	uiPositionXHigh : UINT; // Координаты из того же завершённого FC03-снимка
	uiPositionXLow  : UINT;
	uiPositionYHigh : UINT;
	uiPositionYLow  : UINT;
	uiPositionZHigh : UINT;
	uiPositionZLow  : UINT;
	uiPlcHeartbeat : UINT;
	uiLastRobotHeartbeat : UINT;
	uiCommandCode  : UINT;
	uiRegisterIndex : UINT;
	dwPositionRaw  : DWORD;
	diPositionRaw  : DINT;
	udiReplyTimeoutUs : UDINT;
END_VAR
VAR CONSTANT
	COMMAND_START_ITEM : UINT := UINT#1000; // Документный 1001
	STATUS_START_ITEM  : UINT := UINT#1100; // Документный 1101
	COMMAND_QUANTITY   : UINT := UINT#9;
	STATUS_QUANTITY    : UINT := UINT#17;
	PROTOCOL_VERSION   : UINT := UINT#3;
	RESET_ATTEMPT_TIMEOUT : TIME := T#10S; // Полная попытка: запись, feedback, снятие
	STATUS_CONTROLLER_ON  : UINT := UINT#16#0001;
	STATUS_AUTOMATIC_MODE : UINT := UINT#16#0002;
	STATUS_REMOTE_ENABLED : UINT := UINT#16#0004;
	STATUS_DRIVES_ENABLED : UINT := UINT#16#0008;
	STATUS_HOMED          : UINT := UINT#16#0010;
	STATUS_EMERGENCY_STOP : UINT := UINT#16#0020;
	STATUS_ROBOT_ALARM    : UINT := UINT#16#0040;
	STATUS_ROBOT_READY    : UINT := UINT#16#0080;
	STATUS_POSITION_VALID : UINT := UINT#16#0100;
	STATUS_SIMULATOR_ACTIVE : UINT := UINT#16#0200;
END_VAR

// --- BEGIN IMPLEMENTATION ---

Status.xConfigValid := (Config.aIpAddress[0] > BYTE#0)
	AND (Config.aIpAddress[0] < BYTE#224)
	AND (Config.uiPort > UINT#0)
	AND (Config.uiUnitId <= UINT#255)
	AND (Config.tResponseTimeout >= T#50MS)
	AND (Config.tPollInterval >= T#10MS)
	AND (Config.tHeartbeatTimeout >= T#500MS)
	AND (Config.tCommandTimeout >= T#1S);

	udiReplyTimeoutUs := TIME_TO_UDINT(Config.tResponseTimeout) * UDINT#1000;
	rtStop(CLK := Command.xStop);
	rtReset(CLK := Command.xReset);
	rtReconnect(CLK := xReconnect);
	IF rtStop.Q THEN
		xStopPending := TRUE;
	END_IF;
	IF rtReset.Q AND NOT xResetInProgress THEN
		xResetPending := TRUE;
		xResetInProgress := TRUE;
		xResetWriteDone := FALSE;
		Status.xResetDone := FALSE;
		Status.xResetFailed := FALSE;
	END_IF;
xReadExecute := FALSE;
xWriteExecute := FALSE;
xHeartbeatChanged := FALSE;

fbClient(
	xConnect := xConnect,
	aIPaddr := Config.aIpAddress,
	uiPort := Config.uiPort,
	tConnnectTimeOut := Config.tHeartbeatTimeout
);

IF NOT xEnable OR NOT Status.xConfigValid THEN
	xConnect := FALSE;
	eState := E_ROBOT_MODBUS_CLIENT_STATE.DISABLED;
	xStatusFresh := FALSE;
	xCommandArmed := FALSE;
	xCommandActive := FALSE;
	xWritePending := FALSE;
	xStopPending := FALSE;
	xResetPending := FALSE;
	xResetInProgress := FALSE;
	xResetWriteDone := FALSE;
	Status.xResetDone := FALSE;
	Status.xResetFailed := FALSE;
	xControlClearPending := FALSE;
	xHeartbeatSeen := FALSE;
	xPlcHeartbeatDue := FALSE;
	uiActiveSeq := UINT#0;
	Status.xConnected := FALSE;
ELSE
	xConnect := TRUE;
	IF rtReconnect.Q THEN
		xConnect := FALSE;
		eState := E_ROBOT_MODBUS_CLIENT_STATE.RECONNECT_WAIT;
		xStatusFresh := FALSE;
		xCommandArmed := FALSE;
		xCommandActive := FALSE;
		xWritePending := FALSE;
		xControlClearPending := FALSE;
		xHeartbeatSeen := FALSE;
		xPlcHeartbeatDue := FALSE;
	END_IF;
END_IF;

CASE eState OF
	E_ROBOT_MODBUS_CLIENT_STATE.DISABLED:
		IF xEnable AND Status.xConfigValid THEN
			xConnect := TRUE;
			eState := E_ROBOT_MODBUS_CLIENT_STATE.CONNECTING;
		END_IF;

	E_ROBOT_MODBUS_CLIENT_STATE.CONNECTING:
		IF fbClient.xConnected THEN
			eState := E_ROBOT_MODBUS_CLIENT_STATE.INITIAL_READ;
		ELSIF fbClient.xError THEN
			Status.udiClientError := TO_UDINT(fbClient.eErrorID);
			xConnect := FALSE;
			eState := E_ROBOT_MODBUS_CLIENT_STATE.RECONNECT_WAIT;
		END_IF;

	E_ROBOT_MODBUS_CLIENT_STATE.INITIAL_READ:
		xReadExecute := TRUE;
		IF fbRead.xDone THEN
			xStatusFresh := TRUE;
			uiCommandSeq := auiReadRegisters[0];
			uiActiveSeq := UINT#0;
			uiPlcHeartbeat := UINT#0;
			uiLastRobotHeartbeat := auiReadRegisters[6];
			xHeartbeatSeen := FALSE;
			FOR uiRegisterIndex := UINT#0 TO UINT#8 DO
				auiWriteRegisters[uiRegisterIndex] := UINT#0;
			END_FOR;
			auiWriteRegisters[7] := uiCommandSeq;
			eState := E_ROBOT_MODBUS_CLIENT_STATE.INITIAL_READ_RELEASE;
		ELSIF fbRead.xError THEN
			Status.udiReadError := TO_UDINT(fbRead.eErrorID);
			xConnect := FALSE;
			eState := E_ROBOT_MODBUS_CLIENT_STATE.RECONNECT_WAIT;
		END_IF;

	E_ROBOT_MODBUS_CLIENT_STATE.INITIAL_READ_RELEASE:
		IF NOT fbRead.xBusy THEN
			eState := E_ROBOT_MODBUS_CLIENT_STATE.CLEAR_COMMAND;
		END_IF;

	E_ROBOT_MODBUS_CLIENT_STATE.CLEAR_COMMAND:
		xWriteExecute := TRUE;
		IF fbWrite.xDone THEN
			eState := E_ROBOT_MODBUS_CLIENT_STATE.CLEAR_COMMAND_RELEASE;
		ELSIF fbWrite.xError THEN
			Status.udiWriteError := TO_UDINT(fbWrite.eErrorID);
			xConnect := FALSE;
			eState := E_ROBOT_MODBUS_CLIENT_STATE.RECONNECT_WAIT;
		END_IF;

	E_ROBOT_MODBUS_CLIENT_STATE.CLEAR_COMMAND_RELEASE:
		IF NOT fbWrite.xBusy THEN
			xCommandArmed := NOT Command.xExecute;
			xCommandActive := FALSE;
			eState := E_ROBOT_MODBUS_CLIENT_STATE.READY;
		END_IF;

	E_ROBOT_MODBUS_CLIENT_STATE.READY:
		IF NOT fbClient.xConnected OR fbClient.xError THEN
			Status.udiClientError := TO_UDINT(fbClient.eErrorID);
			xConnect := FALSE;
			eState := E_ROBOT_MODBUS_CLIENT_STATE.RECONNECT_WAIT;
		ELSIF xStopPending THEN
			// Stop отменяет текущую попытку сброса; он не может быть проглочен Reset.
			IF xResetInProgress THEN Status.xResetFailed := TRUE; END_IF;
			xResetInProgress := FALSE;
			xResetWriteDone := FALSE;
			// Stop always preempts Reset and normal commands.
			// Execute снимается сразу: после принятого CommandSeq это не отменяет
			// команду, зато позволяет роботу выйти из DONE/ERROR/STOPPED в IDLE.
			// Без этого уже завершённая дискретная команда навечно удерживала
			// Execute=1, а xControlClearPending ждал недостижимый IDLE.
			auiWriteRegisters[0] := UINT#0;
			auiWriteRegisters[1] := UINT#0;
			auiWriteRegisters[2] := UINT#1;
			auiWriteRegisters[3] := UINT#0;
			auiWriteRegisters[4] := UINT#0;
			auiWriteRegisters[5] := UINT#0;
			auiWriteRegisters[6] := UINT#0;
			xStopPending := FALSE;
			xResetPending := FALSE;
			xControlClearPending := TRUE;
			xWritePending := TRUE;
		ELSIF xResetPending THEN
			// Reset обязан прервать незавершённую очистку Stop. Иначе
			// xControlClearPending имеет приоритет и защёлкнутый Reset никогда
			// не попадает в регистр 1004.
			auiWriteRegisters[0] := UINT#0;
			auiWriteRegisters[1] := UINT#0;
			auiWriteRegisters[2] := UINT#0;
			auiWriteRegisters[3] := UINT#1;
			auiWriteRegisters[4] := UINT#0;
			auiWriteRegisters[5] := UINT#0;
			auiWriteRegisters[6] := UINT#0;
			xCommandActive := FALSE;
			uiActiveSeq := UINT#0;
			xCommandArmed := FALSE;
			xResetPending := FALSE;
			xControlClearPending := TRUE;
			xWritePending := TRUE;
		ELSIF xControlClearPending THEN
			// Stop удерживается до STOPPED/IDLE, Reset — до снятия аварии. Так
			// импульс не потеряется между более медленными циклами программы робота.
			IF ((auiWriteRegisters[2] = UINT#1)
				AND ((Status.uiExecutionState = TO_UINT(E_ROBOT_MODBUS_EXECUTION_STATE.STOPPED))
					OR (Status.uiExecutionState = TO_UINT(E_ROBOT_MODBUS_EXECUTION_STATE.IDLE))))
			OR ((auiWriteRegisters[3] = UINT#1)
				AND xResetWriteDone
				AND NOT Status.xRobotAlarm
				AND (Status.uiExecutionState =
					TO_UINT(E_ROBOT_MODBUS_EXECUTION_STATE.IDLE))) THEN
				auiWriteRegisters[2] := UINT#0;
				auiWriteRegisters[3] := UINT#0;
				xCommandActive := FALSE;
				uiActiveSeq := UINT#0;
				// Верхний FB удерживает Execute до появления Busy. Поэтому после
				// подтверждённой очистки принимаем уже удерживаемую новую команду,
				// а не требуем ещё одного фронта от HMI.
				xCommandArmed := TRUE;
				xControlClearPending := FALSE;
				xWritePending := TRUE;
			END_IF;
		ELSIF Command.xExecute AND xCommandArmed AND NOT xCommandActive THEN
			uiCommandCode := UINT#0;
			CASE Command.eAction OF
				E_ROBOT_ACTION.MOVE_TO_POINT:
					CASE Command.eSetPoint OF
						E_POINT_NAME.MACHINE_1_ABOVE: uiCommandCode := UINT#10;
						E_POINT_NAME.MACHINE_1_INSIDE: uiCommandCode := UINT#11;
						E_POINT_NAME.MACHINE_1_CHUCK_APROACH: uiCommandCode := UINT#12;
						E_POINT_NAME.MACHINE_1_CHUCK_POSITION: uiCommandCode := UINT#13;
						E_POINT_NAME.MACHINE_2_ABOVE: uiCommandCode := UINT#14;
						E_POINT_NAME.MACHINE_2_INSIDE: uiCommandCode := UINT#15;
						E_POINT_NAME.MACHINE_2_CHUCK_APROACH: uiCommandCode := UINT#16;
						E_POINT_NAME.MACHINE_2_CHUCK_POSITION: uiCommandCode := UINT#17;
						E_POINT_NAME.MACHINE_3_ABOVE: uiCommandCode := UINT#18;
						E_POINT_NAME.MACHINE_3_INSIDE: uiCommandCode := UINT#19;
						E_POINT_NAME.MACHINE_3_CHUCK_APROACH: uiCommandCode := UINT#20;
						E_POINT_NAME.MACHINE_3_CHUCK_POSITION: uiCommandCode := UINT#21;
						E_POINT_NAME.HOME_SAFETY: uiCommandCode := UINT#22;
						E_POINT_NAME.MAGAZINE_SAFE: uiCommandCode := UINT#23;
						E_POINT_NAME.MAGAZINE_CHANGE: uiCommandCode := UINT#24;
						E_POINT_NAME.MAGAZINE_IN_SLOT: uiCommandCode := UINT#25;
					END_CASE;
				E_ROBOT_ACTION.UNCLAMP_1: uiCommandCode := UINT#2;
				E_ROBOT_ACTION.CLAMP_1: uiCommandCode := UINT#3;
				E_ROBOT_ACTION.UNCLAMP_2: uiCommandCode := UINT#4;
				E_ROBOT_ACTION.CLAMP_2: uiCommandCode := UINT#5;
				E_ROBOT_ACTION.ROTATE_TO_BLANK: uiCommandCode := UINT#6;
				E_ROBOT_ACTION.ROTATE_TO_DETAIL: uiCommandCode := UINT#7;
			END_CASE;

			IF uiCommandCode > UINT#0 THEN
				uiCommandSeq := uiCommandSeq + UINT#1;
				IF uiCommandSeq = UINT#0 THEN
					uiCommandSeq := UINT#1;
				END_IF;
				uiActiveSeq := uiCommandSeq;
				auiWriteRegisters[0] := uiCommandCode;
				auiWriteRegisters[1] := UINT#1;
				auiWriteRegisters[2] := UINT#0;
				auiWriteRegisters[3] := UINT#0;
				auiWriteRegisters[4] := SINT_TO_UINT(Command.iActiveSlot);
				auiWriteRegisters[5] := Command.uiMagazineId;
				auiWriteRegisters[6] := UINT#0;
				auiWriteRegisters[7] := uiCommandSeq;
				xCommandActive := TRUE;
				xCommandArmed := FALSE;
				xWritePending := TRUE;
			END_IF;
		ELSIF NOT Command.xExecute AND xCommandActive THEN
			auiWriteRegisters[0] := UINT#0;
			auiWriteRegisters[1] := UINT#0;
			auiWriteRegisters[2] := UINT#0;
			auiWriteRegisters[3] := UINT#0;
			auiWriteRegisters[4] := UINT#0;
			auiWriteRegisters[5] := UINT#0;
			auiWriteRegisters[6] := UINT#0;
			xCommandActive := FALSE;
			// CommandSeq в регистре сохраняется как последний использованный номер,
			// но завершённая транзакция больше не имеет права публиковать Done.
			// Повтор после Reset всегда получит новый ненулевой sequence.
			uiActiveSeq := UINT#0;
			xCommandArmed := TRUE;
			xWritePending := TRUE;
		ELSIF NOT Command.xExecute THEN
			xCommandArmed := TRUE;
		END_IF;

		IF xPlcHeartbeatDue THEN
			uiPlcHeartbeat := uiPlcHeartbeat + UINT#1;
			auiWriteRegisters[8] := uiPlcHeartbeat;
			xPlcHeartbeatDue := FALSE;
			xWritePending := TRUE;
		END_IF;

		IF xWritePending THEN
			eState := E_ROBOT_MODBUS_CLIENT_STATE.WRITE_COMMAND;
		ELSIF tonPoll.Q THEN
			eState := E_ROBOT_MODBUS_CLIENT_STATE.READ_STATUS;
		END_IF;

	E_ROBOT_MODBUS_CLIENT_STATE.WRITE_COMMAND:
		xWriteExecute := TRUE;
		IF fbWrite.xDone THEN
			IF xResetInProgress THEN
				IF auiWriteRegisters[3] = UINT#1 THEN
					xResetWriteDone := TRUE;
				ELSIF xResetWriteDone AND NOT xControlClearPending THEN
					// Успех только после FC03 без аварии/с IDLE и последующей
					// подтверждённой записи Reset=0. Один локальный скан не Ack.
					xResetInProgress := FALSE;
					Status.xResetDone := TRUE;
				END_IF;
			END_IF;
			xWritePending := FALSE;
			eState := E_ROBOT_MODBUS_CLIENT_STATE.WRITE_COMMAND_RELEASE;
		ELSIF fbWrite.xError THEN
			Status.udiWriteError := TO_UDINT(fbWrite.eErrorID);
			xConnect := FALSE;
			eState := E_ROBOT_MODBUS_CLIENT_STATE.RECONNECT_WAIT;
		END_IF;

	E_ROBOT_MODBUS_CLIENT_STATE.WRITE_COMMAND_RELEASE:
		IF NOT fbWrite.xBusy THEN
			eState := E_ROBOT_MODBUS_CLIENT_STATE.READ_STATUS;
		END_IF;

	E_ROBOT_MODBUS_CLIENT_STATE.READ_STATUS:
		xReadExecute := TRUE;
		IF fbRead.xDone THEN
			xStatusFresh := TRUE;
			eState := E_ROBOT_MODBUS_CLIENT_STATE.READ_STATUS_RELEASE;
		ELSIF fbRead.xError THEN
			Status.udiReadError := TO_UDINT(fbRead.eErrorID);
			xConnect := FALSE;
			eState := E_ROBOT_MODBUS_CLIENT_STATE.RECONNECT_WAIT;
		END_IF;

	E_ROBOT_MODBUS_CLIENT_STATE.READ_STATUS_RELEASE:
		IF NOT fbRead.xBusy THEN
			eState := E_ROBOT_MODBUS_CLIENT_STATE.READY;
		END_IF;

	E_ROBOT_MODBUS_CLIENT_STATE.RECONNECT_WAIT:
		xConnect := FALSE;
		xStatusFresh := FALSE;
		IF tonReconnect.Q THEN
			xConnect := TRUE;
			eState := E_ROBOT_MODBUS_CLIENT_STATE.CONNECTING;
		END_IF;
END_CASE;

tonResetAttempt(IN := xResetInProgress, PT := RESET_ATTEMPT_TIMEOUT);
IF xResetInProgress
AND ((eState = E_ROBOT_MODBUS_CLIENT_STATE.RECONNECT_WAIT)
	OR rtReconnect.Q OR tonResetAttempt.Q OR NOT Command.xReset) THEN
	// Не повторяем неоднозначную запись после обрыва. Reconnect сначала
	// прочитает состояние и очистит блок; новый Reset требует нового фронта.
	xResetInProgress := FALSE;
	xResetPending := FALSE;
	xResetWriteDone := FALSE;
	Status.xResetDone := FALSE;
	Status.xResetFailed := TRUE;
	xConnect := FALSE;
	xStatusFresh := FALSE;
	eState := E_ROBOT_MODBUS_CLIENT_STATE.RECONNECT_WAIT;
END_IF;
IF eState = E_ROBOT_MODBUS_CLIENT_STATE.RECONNECT_WAIT THEN
	xReadExecute := FALSE;
	xWriteExecute := FALSE;
	xControlClearPending := FALSE;
	xWritePending := FALSE;
	xCommandArmed := FALSE;
END_IF;
Status.xResetBusy := xResetInProgress;

fbRead(
	xExecute := xReadExecute,
	udiTimeOut := udiReplyTimeoutUs,
	rClient := fbClient,
	uiUnitId := Config.uiUnitId,
	udiReplyTimeout := udiReplyTimeoutUs,
	uiMaxRetries := UINT#1,
	uiStartItem := STATUS_START_ITEM,
	uiQuantity := STATUS_QUANTITY,
	pData := ADR(auiReadRegisters)
);
fbWrite(
	xExecute := xWriteExecute,
	udiTimeOut := udiReplyTimeoutUs,
	rClient := fbClient,
	uiUnitId := Config.uiUnitId,
	udiReplyTimeout := udiReplyTimeoutUs,
	uiMaxRetries := UINT#1,
	uiStartItem := COMMAND_START_ITEM,
	uiQuantity := COMMAND_QUANTITY,
	pData := ADR(auiWriteRegisters)
);

// FC03 может завершиться внутри вызова fbRead. Декодирование выполняется после
// вызова, чтобы технологический Status и сырые диагностические регистры всегда
// относились к одному и тому же снимку опроса.
IF fbRead.xDone THEN
	Status.uiAckSeq := auiReadRegisters[0];
	Status.uiExecutionState := auiReadRegisters[1];
	Status.uiResultCode := auiReadRegisters[2];
	Status.uiActiveCommand := auiReadRegisters[3];
	Status.uiCurrentPoint := auiReadRegisters[4];
	Status.uiGripperStatus := auiReadRegisters[5];
	Status.uiRobotHeartbeat := auiReadRegisters[6];
	Status.uiStatusWord := auiReadRegisters[7];
	Status.uiAlarmCode := auiReadRegisters[8];
	Status.uiOperationPhase := auiReadRegisters[15];
	Status.uiProtocolVersion := auiReadRegisters[16];
	uiDecodedRobotHeartbeat := auiReadRegisters[6];
	uiPositionXHigh := auiReadRegisters[9];
	uiPositionXLow := auiReadRegisters[10];
	uiPositionYHigh := auiReadRegisters[11];
	uiPositionYLow := auiReadRegisters[12];
	uiPositionZHigh := auiReadRegisters[13];
	uiPositionZLow := auiReadRegisters[14];
END_IF;

tonPoll(IN := eState = E_ROBOT_MODBUS_CLIENT_STATE.READY, PT := Config.tPollInterval);
// Heartbeat timer is independent of request states. The due latch prevents a pulse
// from being lost while FC03/FC16 is busy.
tonPlcHeartbeat(
	IN := xEnable AND fbClient.xConnected AND NOT tonPlcHeartbeat.Q,
	PT := T#100MS
);
IF tonPlcHeartbeat.Q THEN
	xPlcHeartbeatDue := TRUE;
END_IF;
tonReconnect(IN := eState = E_ROBOT_MODBUS_CLIENT_STATE.RECONNECT_WAIT, PT := T#1S);

Status.xConnected := fbClient.xConnected AND xConnect;
Status.xStatusFresh := xStatusFresh;

IF uiDecodedRobotHeartbeat <> uiLastRobotHeartbeat THEN
	uiLastRobotHeartbeat := uiDecodedRobotHeartbeat;
	xHeartbeatChanged := TRUE;
	xHeartbeatSeen := TRUE;
END_IF;
tonRobotHeartbeat(
	IN := xEnable AND xStatusFresh AND NOT xHeartbeatChanged,
	PT := Config.tHeartbeatTimeout
);
Status.xCommunicationAlive := Status.xConnected
	AND xStatusFresh
	AND xHeartbeatSeen
	AND NOT tonRobotHeartbeat.Q
	AND (Status.uiProtocolVersion = PROTOCOL_VERSION);
tonCommunicationGrace(
	IN := xEnable AND Status.xConfigValid AND NOT Status.xCommunicationAlive,
	PT := Config.tHeartbeatTimeout
);

Status.xControllerOn := (Status.uiStatusWord AND STATUS_CONTROLLER_ON) <> UINT#0;
Status.xAutomaticMode := (Status.uiStatusWord AND STATUS_AUTOMATIC_MODE) <> UINT#0;
Status.xRemoteEnabled := (Status.uiStatusWord AND STATUS_REMOTE_ENABLED) <> UINT#0;
Status.xDrivesEnabled := (Status.uiStatusWord AND STATUS_DRIVES_ENABLED) <> UINT#0;
Status.xHomed := (Status.uiStatusWord AND STATUS_HOMED) <> UINT#0;
Status.xEmergencyStop := (Status.uiStatusWord AND STATUS_EMERGENCY_STOP) <> UINT#0;
Status.xRobotAlarm := ((Status.uiStatusWord AND STATUS_ROBOT_ALARM) <> UINT#0)
	OR (Status.uiAlarmCode <> UINT#0);
Status.xPositionValid := (Status.uiStatusWord AND STATUS_POSITION_VALID) <> UINT#0;
Status.xSimulatorActive := (Status.uiStatusWord AND STATUS_SIMULATOR_ACTIVE) <> UINT#0;
Status.xReady := Status.xCommunicationAlive
	AND Status.xControllerOn
	AND Status.xAutomaticMode
	AND Status.xRemoteEnabled
	AND Status.xDrivesEnabled
	AND Status.xHomed
	AND Status.xPositionValid
	AND NOT Status.xEmergencyStop
	AND NOT Status.xRobotAlarm
	AND ((Status.uiStatusWord AND STATUS_ROBOT_READY) <> UINT#0);

Status.xDone := (uiActiveSeq <> UINT#0)
	AND xCommandActive
	AND (Status.uiAckSeq = uiActiveSeq)
	AND (Status.uiExecutionState = TO_UINT(E_ROBOT_MODBUS_EXECUTION_STATE.DONE))
	AND (Status.uiResultCode = UINT#0);
// Busy означает активную PLC-транзакцию, включая ожидание AckSeq. Благодаря
// этому FB_ROBOT обязательно увидит запуск новой команды до её terminal state.
Status.xBusy := (uiActiveSeq <> UINT#0)
	AND xCommandActive
	AND NOT Status.xDone
	AND NOT ((Status.uiAckSeq = uiActiveSeq)
		AND ((Status.uiExecutionState = TO_UINT(E_ROBOT_MODBUS_EXECUTION_STATE.ERROR))
			OR (Status.uiExecutionState = TO_UINT(E_ROBOT_MODBUS_EXECUTION_STATE.STOPPED))
			OR ((Status.uiExecutionState = TO_UINT(E_ROBOT_MODBUS_EXECUTION_STATE.DONE))
				AND (Status.uiResultCode <> UINT#0))));
tonCommandTimeout(
	IN := xCommandActive AND NOT Status.xDone,
	PT := Config.tCommandTimeout
);
Status.xCommandTimeout := tonCommandTimeout.Q;
Status.xError := tonCommunicationGrace.Q
	OR Status.xResetFailed
	OR Status.xRobotAlarm
	OR Status.xCommandTimeout
	OR ((uiActiveSeq <> UINT#0)
		AND (Status.uiAckSeq = uiActiveSeq)
		AND ((Status.uiExecutionState = TO_UINT(E_ROBOT_MODBUS_EXECUTION_STATE.ERROR))
			OR ((Status.uiExecutionState = TO_UINT(E_ROBOT_MODBUS_EXECUTION_STATE.DONE))
				AND (Status.uiResultCode <> UINT#0))));

dwPositionRaw := SHL(UINT_TO_DWORD(uiPositionXHigh), 16)
	OR UINT_TO_DWORD(uiPositionXLow);
diPositionRaw := DWORD_TO_DINT(dwPositionRaw);
Status.lrActualX := DINT_TO_LREAL(diPositionRaw) / LREAL#10.0;
dwPositionRaw := SHL(UINT_TO_DWORD(uiPositionYHigh), 16)
	OR UINT_TO_DWORD(uiPositionYLow);
diPositionRaw := DWORD_TO_DINT(dwPositionRaw);
Status.lrActualY := DINT_TO_LREAL(diPositionRaw) / LREAL#10.0;
dwPositionRaw := SHL(UINT_TO_DWORD(uiPositionZHigh), 16)
	OR UINT_TO_DWORD(uiPositionZLow);
diPositionRaw := DWORD_TO_DINT(dwPositionRaw);
Status.lrActualZ := DINT_TO_LREAL(diPositionRaw) / LREAL#10.0;

(* ---- FB_SIMULATION_DYNAMIC_LIMITS.st ---- *)
FUNCTION_BLOCK FB_SIMULATION_DYNAMIC_LIMITS
VAR_INPUT
	xSimulationMode : BOOL; // Активна тестовая среда SIMULATION
	xSoftMotionMode : BOOL; // Роботом управляют локальные оси SoftMotion
	xAccelerationEnabled : BOOL; // Для следующего теста выбран ускоренный профиль
	xPrepareTest : BOOL; // Фронт подготовки следующего сценария
	uiRequestedFactor : UINT; // Запрошенное масштабирование времени 1..100
	xCellRunning : BOOL;
	xRobotBusy : BOOL;
	xMotionBusy : BOOL;
	xDrivesPowered : BOOL;
	xDrivesOff : BOOL;
	eGroupState : E_AXIS_GROUP_STATE;
	tTransactionTimeout : TIME := T#60S; // Общий предел Stop -> Disable -> Change -> Enable
END_VAR
VAR_OUTPUT
	xCellStopRequest : BOOL; // Сначала остановить технологический цикл
	xMotionStopRequest : BOOL; // Затем остановить движение группы
	xGroupDisableRequest : BOOL; // Перед изменением лимитов получить GroupDisabled
	xDrivesEnableRequest : BOOL; // После изменения вернуть штатную готовность
	xBusy : BOOL;
	xPending : BOOL; // Ползунок изменён; значение ждёт границы следующего теста
	xReadyForTest : BOOL; // Новый тест можно запускать
	xAccelerationActive : BOOL;
	uiAppliedFactor : UINT := UINT#1;
	xDone : BOOL;
	xError : BOOL;
	udiErrorId : UDINT;
END_VAR
VAR_IN_OUT
	AxisX : AXIS_REF_SM3;
	AxisY : AXIS_REF_SM3;
	AxisZ : AXIS_REF_SM3;
END_VAR
VAR CONSTANT
	STATE_IDLE : UINT := UINT#0;
	STATE_WAIT_STANDSTILL : UINT := UINT#10;
	STATE_WAIT_GROUP_DISABLED : UINT := UINT#20;
	STATE_CHANGE_X : UINT := UINT#30;
	STATE_CHANGE_Y : UINT := UINT#40;
	STATE_CHANGE_Z : UINT := UINT#50;
	STATE_PREPARE_ROLLBACK : UINT := UINT#55;
	STATE_WAIT_REENABLE : UINT := UINT#60;
	STATE_LOCKED_ERROR : UINT := UINT#90;
	ERR_INVALID_ORIGINAL_LIMITS : UDINT := UDINT#16#80010001;
	ERR_TRANSACTION_TIMEOUT : UDINT := UDINT#16#80010002;
	ERR_INVALID_STATE : UDINT := UDINT#16#80010003;
END_VAR
VAR
	rtPrepareTest : R_TRIG;
	tonTransaction : TON;
	uiState : UINT := UINT#0;
	uiAxis : UINT;
	uiDesiredFactor : UINT := UINT#1;
	uiTargetFactor : UINT := UINT#1;
	xOriginalLimitsSaved : BOOL;
	xOriginalLimitsValid : BOOL;
	xRestoreOnExit : BOOL;
	xRollback : BOOL;
	xReenableAfterChange : BOOL;

	alrOriginalVelocity : ARRAY [1..3] OF LREAL;
	alrOriginalAcceleration : ARRAY [1..3] OF LREAL;
	alrOriginalDeceleration : ARRAY [1..3] OF LREAL;
	alrOriginalJerk : ARRAY [1..3] OF LREAL;
	alrTargetVelocity : ARRAY [1..3] OF LREAL;
	alrTargetAcceleration : ARRAY [1..3] OF LREAL;
	alrTargetDeceleration : ARRAY [1..3] OF LREAL;
	alrTargetJerk : ARRAY [1..3] OF LREAL;
	lrFactor : LREAL;
	lrFactorSquared : LREAL;
	lrFactorCubed : LREAL;

	fbChangeX : SMC_ChangeDynamicLimits;
	fbChangeY : SMC_ChangeDynamicLimits;
	fbChangeZ : SMC_ChangeDynamicLimits;
END_VAR

// --- BEGIN IMPLEMENTATION ---

// Запрошенное значение разрешено менять когда угодно. Оно только создаёт
// pending-запрос; уже выполняемая траектория никогда не перепланируется.
uiDesiredFactor := MAX(UINT#1, MIN(UINT#100, uiRequestedFactor));
IF NOT (xSimulationMode AND xSoftMotionMode AND xAccelerationEnabled) THEN
	uiDesiredFactor := UINT#1;
END_IF;
rtPrepareTest(CLK := xPrepareTest);

xCellStopRequest := FALSE;
xMotionStopRequest := FALSE;
xGroupDisableRequest := FALSE;
xDrivesEnableRequest := FALSE;
xDone := FALSE;

// Штатные лимиты снимаются ровно при входе в SoftMotion-симуляцию, до первого
// масштабирования. Прямое редактирование AXIS_REF здесь не выполняется.
IF xSimulationMode AND xSoftMotionMode AND NOT xOriginalLimitsSaved THEN
	// Dynamic limits из конфигуратора оси находятся в fSWMax*. fMax* — это
	// remote limits самого привода и у виртуальной оси законно остаются нулями.
	alrOriginalVelocity[1] := AxisX.fSWMaxVelocity;
	alrOriginalAcceleration[1] := AxisX.fSWMaxAcceleration;
	alrOriginalDeceleration[1] := AxisX.fSWMaxDeceleration;
	alrOriginalJerk[1] := AxisX.fSWMaxJerk;
	alrOriginalVelocity[2] := AxisY.fSWMaxVelocity;
	alrOriginalAcceleration[2] := AxisY.fSWMaxAcceleration;
	alrOriginalDeceleration[2] := AxisY.fSWMaxDeceleration;
	alrOriginalJerk[2] := AxisY.fSWMaxJerk;
	alrOriginalVelocity[3] := AxisZ.fSWMaxVelocity;
	alrOriginalAcceleration[3] := AxisZ.fSWMaxAcceleration;
	alrOriginalDeceleration[3] := AxisZ.fSWMaxDeceleration;
	alrOriginalJerk[3] := AxisZ.fSWMaxJerk;

	IF alrOriginalVelocity[1] <= LREAL#0.0 THEN alrOriginalVelocity[1] := AxisX.fMaxVelocity; END_IF;
	IF alrOriginalAcceleration[1] <= LREAL#0.0 THEN alrOriginalAcceleration[1] := AxisX.fMaxAcceleration; END_IF;
	IF alrOriginalDeceleration[1] <= LREAL#0.0 THEN alrOriginalDeceleration[1] := AxisX.fMaxDeceleration; END_IF;
	IF alrOriginalJerk[1] <= LREAL#0.0 THEN alrOriginalJerk[1] := AxisX.fMaxJerk; END_IF;
	IF alrOriginalVelocity[2] <= LREAL#0.0 THEN alrOriginalVelocity[2] := AxisY.fMaxVelocity; END_IF;
	IF alrOriginalAcceleration[2] <= LREAL#0.0 THEN alrOriginalAcceleration[2] := AxisY.fMaxAcceleration; END_IF;
	IF alrOriginalDeceleration[2] <= LREAL#0.0 THEN alrOriginalDeceleration[2] := AxisY.fMaxDeceleration; END_IF;
	IF alrOriginalJerk[2] <= LREAL#0.0 THEN alrOriginalJerk[2] := AxisY.fMaxJerk; END_IF;
	IF alrOriginalVelocity[3] <= LREAL#0.0 THEN alrOriginalVelocity[3] := AxisZ.fMaxVelocity; END_IF;
	IF alrOriginalAcceleration[3] <= LREAL#0.0 THEN alrOriginalAcceleration[3] := AxisZ.fMaxAcceleration; END_IF;
	IF alrOriginalDeceleration[3] <= LREAL#0.0 THEN alrOriginalDeceleration[3] := AxisZ.fMaxDeceleration; END_IF;
	IF alrOriginalJerk[3] <= LREAL#0.0 THEN alrOriginalJerk[3] := AxisZ.fMaxJerk; END_IF;

	xOriginalLimitsValid := TRUE;
	FOR uiAxis := UINT#1 TO UINT#3 DO
		xOriginalLimitsValid := xOriginalLimitsValid
			AND (alrOriginalVelocity[uiAxis] > LREAL#0.0)
			AND (alrOriginalAcceleration[uiAxis] > LREAL#0.0)
			AND (alrOriginalDeceleration[uiAxis] > LREAL#0.0)
			AND (alrOriginalJerk[uiAxis] > LREAL#0.0);
	END_FOR;
	IF xOriginalLimitsValid THEN
		xOriginalLimitsSaved := TRUE;
		uiAppliedFactor := UINT#1;
		xError := FALSE;
		udiErrorId := UDINT#0;
	ELSIF rtPrepareTest.Q THEN
		// До подготовки теста просто ждём инициализацию осей; не защёлкиваем
		// ложную ошибку на первом цикле после переключения среды.
		xError := TRUE;
		udiErrorId := ERR_INVALID_ORIGINAL_LIMITS;
	END_IF;
END_IF;

// Ошибка чтения исходных лимитов не должна блокировать обычную ячейку после
// выхода из тестовой среды и не должна переживать Online Change этого исправления.
IF NOT xSimulationMode
AND NOT xOriginalLimitsSaved
AND (uiState = STATE_IDLE)
AND (udiErrorId = ERR_INVALID_ORIGINAL_LIMITS) THEN
	xError := FALSE;
	udiErrorId := UDINT#0;
END_IF;

xRestoreOnExit := xOriginalLimitsSaved
	AND (NOT xSimulationMode OR NOT xSoftMotionMode)
	AND (uiAppliedFactor <> UINT#1);
xPending := xOriginalLimitsSaved AND (uiDesiredFactor <> uiAppliedFactor);

// Один общий таймаут защищает всю транзакцию Stop -> Disable -> Change -> Enable.
tonTransaction(IN := uiState <> STATE_IDLE, PT := tTransactionTimeout);
IF tonTransaction.Q
AND (uiState <> STATE_IDLE)
AND (uiState <> STATE_LOCKED_ERROR) THEN
	xError := TRUE;
	udiErrorId := ERR_TRANSACTION_TIMEOUT;
	uiState := STATE_LOCKED_ERROR;
END_IF;

CASE uiState OF
	STATE_IDLE:
		xBusy := FALSE;
		// Возврат штатных лимитов при выходе из SIMULATION выполняется сразу.
		// Обычная ячейка не получит Start, пока транзакция не закончена.
		IF xRestoreOnExit THEN
			xError := FALSE;
			udiErrorId := UDINT#0;
			uiTargetFactor := UINT#1;
			xRollback := FALSE;
			xReenableAfterChange := xSoftMotionMode AND NOT xDrivesOff;
			xBusy := TRUE;
			uiState := STATE_WAIT_STANDSTILL;
		ELSIF rtPrepareTest.Q
		AND xSimulationMode
		AND xSoftMotionMode
		AND xPending
		AND NOT xCellRunning THEN
			xError := FALSE;
			udiErrorId := UDINT#0;
			uiTargetFactor := uiDesiredFactor;
			xRollback := FALSE;
			xReenableAfterChange := NOT xDrivesOff;
			xBusy := TRUE;
			uiState := STATE_WAIT_STANDSTILL;
		ELSIF NOT xSimulationMode
		AND xOriginalLimitsSaved
		AND (uiAppliedFactor = UINT#1) THEN
			// Лимиты не менялись либо уже успешно восстановлены.
			xOriginalLimitsSaved := FALSE;
		END_IF;

	STATE_WAIT_STANDSTILL:
		xBusy := TRUE;
		xCellStopRequest := xCellRunning;
		xMotionStopRequest := xMotionBusy OR xRobotBusy;
		IF NOT xCellRunning AND NOT xMotionBusy AND NOT xRobotBusy THEN
			uiState := STATE_WAIT_GROUP_DISABLED;
		END_IF;

	STATE_WAIT_GROUP_DISABLED:
		xBusy := TRUE;
		xGroupDisableRequest := NOT xDrivesOff;
		IF xDrivesOff AND (eGroupState = E_AXIS_GROUP_STATE.DISABLED) THEN
			IF xRollback THEN
				FOR uiAxis := UINT#1 TO UINT#3 DO
					alrTargetVelocity[uiAxis] := alrOriginalVelocity[uiAxis];
					alrTargetAcceleration[uiAxis] := alrOriginalAcceleration[uiAxis];
					alrTargetDeceleration[uiAxis] := alrOriginalDeceleration[uiAxis];
					alrTargetJerk[uiAxis] := alrOriginalJerk[uiAxis];
				END_FOR;
			ELSE
				lrFactor := UINT_TO_LREAL(uiTargetFactor);
				lrFactorSquared := lrFactor * lrFactor;
				lrFactorCubed := lrFactorSquared * lrFactor;
				alrTargetVelocity[1] := alrOriginalVelocity[1] * lrFactor;
				alrTargetAcceleration[1] := alrOriginalAcceleration[1] * lrFactorSquared;
				alrTargetDeceleration[1] := alrOriginalDeceleration[1] * lrFactorSquared;
				alrTargetJerk[1] := alrOriginalJerk[1] * lrFactorCubed;
				alrTargetVelocity[2] := alrOriginalVelocity[2] * lrFactor;
				alrTargetAcceleration[2] := alrOriginalAcceleration[2] * lrFactorSquared;
				alrTargetDeceleration[2] := alrOriginalDeceleration[2] * lrFactorSquared;
				alrTargetJerk[2] := alrOriginalJerk[2] * lrFactorCubed;
				alrTargetVelocity[3] := alrOriginalVelocity[3] * lrFactor;
				alrTargetAcceleration[3] := alrOriginalAcceleration[3] * lrFactorSquared;
				alrTargetDeceleration[3] := alrOriginalDeceleration[3] * lrFactorSquared;
				alrTargetJerk[3] := alrOriginalJerk[3] * lrFactorCubed;
			END_IF;
			uiState := STATE_CHANGE_X;
		END_IF;

	STATE_CHANGE_X:
		xBusy := TRUE;
		IF fbChangeX.bError THEN
			xError := TRUE;
			udiErrorId := TO_UDINT(fbChangeX.ErrorID);
			IF xRollback THEN uiState := STATE_LOCKED_ERROR;
			ELSE uiState := STATE_PREPARE_ROLLBACK; END_IF;
		ELSIF fbChangeX.bDone THEN
			uiState := STATE_CHANGE_Y;
		END_IF;

	STATE_CHANGE_Y:
		xBusy := TRUE;
		IF fbChangeY.bError THEN
			xError := TRUE;
			udiErrorId := TO_UDINT(fbChangeY.ErrorID);
			IF xRollback THEN uiState := STATE_LOCKED_ERROR;
			ELSE uiState := STATE_PREPARE_ROLLBACK; END_IF;
		ELSIF fbChangeY.bDone THEN
			uiState := STATE_CHANGE_Z;
		END_IF;

	STATE_CHANGE_Z:
		xBusy := TRUE;
		IF fbChangeZ.bError THEN
			xError := TRUE;
			udiErrorId := TO_UDINT(fbChangeZ.ErrorID);
			IF xRollback THEN uiState := STATE_LOCKED_ERROR;
			ELSE uiState := STATE_PREPARE_ROLLBACK; END_IF;
		ELSIF fbChangeZ.bDone THEN
			IF xReenableAfterChange THEN
				uiState := STATE_WAIT_REENABLE;
			ELSE
				IF xRollback THEN uiAppliedFactor := UINT#1;
				ELSE uiAppliedFactor := uiTargetFactor; END_IF;
				xDone := NOT xRollback;
				xBusy := FALSE;
				uiState := STATE_IDLE;
			END_IF;
		END_IF;

	STATE_PREPARE_ROLLBACK:
		// Один цикл с Execute=FALSE создаёт корректный новый фронт для X.
		xBusy := TRUE;
		xRollback := TRUE;
		uiState := STATE_WAIT_GROUP_DISABLED;

	STATE_WAIT_REENABLE:
		xBusy := TRUE;
		xDrivesEnableRequest := TRUE;
		IF xDrivesPowered AND (eGroupState = E_AXIS_GROUP_STATE.READY) THEN
			IF xRollback THEN uiAppliedFactor := UINT#1;
			ELSE uiAppliedFactor := uiTargetFactor; END_IF;
			xDone := NOT xRollback;
			xBusy := FALSE;
			uiState := STATE_IDLE;
		END_IF;

	STATE_LOCKED_ERROR:
		// При неизвестном/неустранимом результате оставляем группу отключённой.
		// Следующий Start заблокирован, пока инженер не устранит причину.
		xBusy := FALSE;
		xGroupDisableRequest := NOT xDrivesOff;

ELSE
	xError := TRUE;
	udiErrorId := ERR_INVALID_STATE;
	uiState := STATE_LOCKED_ERROR;
END_CASE;

fbChangeX(
	Axis := AxisX,
	bExecute := uiState = STATE_CHANGE_X,
	fMaxVelocity := alrTargetVelocity[1],
	fMaxAcceleration := alrTargetAcceleration[1],
	fMaxDeceleration := alrTargetDeceleration[1],
	fMaxJerk := alrTargetJerk[1]
);
fbChangeY(
	Axis := AxisY,
	bExecute := uiState = STATE_CHANGE_Y,
	fMaxVelocity := alrTargetVelocity[2],
	fMaxAcceleration := alrTargetAcceleration[2],
	fMaxDeceleration := alrTargetDeceleration[2],
	fMaxJerk := alrTargetJerk[2]
);
fbChangeZ(
	Axis := AxisZ,
	bExecute := uiState = STATE_CHANGE_Z,
	fMaxVelocity := alrTargetVelocity[3],
	fMaxAcceleration := alrTargetAcceleration[3],
	fMaxDeceleration := alrTargetDeceleration[3],
	fMaxJerk := alrTargetJerk[3]
);

xPending := xOriginalLimitsSaved AND (uiDesiredFactor <> uiAppliedFactor);
xAccelerationActive := xSimulationMode AND xSoftMotionMode
	AND (uiAppliedFactor > UINT#1) AND NOT xError;
xReadyForTest := NOT xBusy AND NOT xError
	AND (NOT (xSimulationMode AND xSoftMotionMode AND xAccelerationEnabled) OR NOT xPending);
